(* CODESYS project RobotLibrary.library
   Company: Thorsten Brach
   Description: SRCI Robot Library
   Version: 1.5.7.0
   Placeholder: RobotLibrary
   Author: Thorsten Brach
   Title: RobotLibrary

Project tree, tasks and I/O mapping:
  libraries: RobotLibrarySysDep, * (Thorsten Brach); Tc2_Standard, 3.4.5.0 (Beckhoff Automation GmbH)
  Library/
    Constants/
      global variables RobotLibraryConstants
      global variables RobotLibraryDefines
    Enumerations/
      ArmConfig/
        data type ArmConfigElbow
        data type ArmConfigShoulder
        data type ArmConfigWrist
      Events/
        data type RobotLibraryErrorIdEnum
        data type RobotLibraryInfoIdEnum
        data type RobotLibraryWarningIdEnum
      Flag/
        data type SequenceFlag
        data type SequenceFlagEnum
      Level/
        data type LogLevel
        data type LogLevelEnum
        data type MessageLevel
        data type MessageLevelEnum
        data type PriorityLevel
      Miscellaneous/
        data type AxisUnit
        data type CircPlane
        data type ComDirection
        data type ControlHalfByte
        data type ErrorReaction
        data type LoadMeasurementSteps
        data type PathChoice
        data type ReferenceElement
        data type Severity
        data type SyncDirection
        data type SyncReaction
        data type SyncTime
        data type TriggerCondition
        data type UnitLimitAxis
      Mode/
        data type AbortingMode
        data type AbortingModeEnum
        data type BlendingMode
        data type CircMode
        data type CollisionReactionMode
        data type ConnectionMode
        data type DefinitionMode
        data type DetectionMode
        data type ErrorTriggerMode
        data type ExecutionMode
        data type FrameCalculationMode
        data type FunctionMode
        data type InterpolationMode
        data type JogMode
        data type LimitMode
        data type LoadMeasurementMode
        data type LogonMode
        data type MeasuringIoMode
        data type MeasuringUnitMode
        data type OperationMode
        data type OrientationMode
        data type OriMode
        data type ProcessingMode
        data type ProcessingModeEnum
        data type ResistanceForceMode
        data type ReturnMode
        data type SensorConnectionMode
        data type SingularityAvoidanceMode
        data type SplineMode
        data type StepMode
        data type StopMode
        data type SyncInMode
        data type SyncMode
        data type ThresholdMode
        data type ToolCalculationMode
        data type TrajectoryMode
        data type TransformMode
        data type TriggerModeIo
        data type TriggerModeLimit
        data type TriggerModeMeasurement
        data type TriggerReactionMode
        data type TurnMode
        data type WorkAreaReactionMode
      State/
        data type ActiveCommandRegisterState
        data type BufferStateCmd
        data type BufferStateRsp
        data type CmdMessageState
        data type InitializationState
        data type RaPowerState
        data type RaSequenceState
        data type RiState
        data type TelegramState
      Type/
        data type AreaType
        data type AreaTypeEnum
        data type AxesGroupParameterCmdEntries
        data type CmdType
        data type ConveyorType
        data type DataType
        data type MessageType
        data type ReferenceType
        data type UnitType
    Functions/
      Check/
        function IsDefaultDynamicsEqual [ST]
        function IsFrameDataEqual [ST]
        function IsLoadDataEqual [ST]
        function IsReferenceDynamicsEqual [ST]
        function IsSwLimitsEqual [ST]
        function IsToolDataEqual [ST]
        function IsWorkAreaEqual [ST]
      Common/
        function CheckTimeout [ST]
        function SetTimeout [ST]
      Convert/
        DT/
          function DATE_TO_IEC_DATE [ST]
          function IEC_DATE_TO_DATE [ST]
          function IEC_TIME_TO_TIME [ST]
          function IEC_TIMESTAMP_TO_DT [ST]
          function IEC_TIMESTAMP_TO_SYSTEMTIME [ST]
          function SYSTEMTIME_TO_IEC_TIMESTAMP [ST]
          function TIME_TO_IEC_TIME [ST]
        Misc/
          function ArmConfigParameterToBytes [ST]
          function BytesToRCSupportedFunctions [ST]
          function ByteToAxisExternalUnit [ST]
          function ByteToAxisExternalUsed [ST]
          function ByteToAxisJointUnit [ST]
          function ByteToAxisJointUsed [ST]
          function ByteToFragmentAction [ST]
          function ByteToVersion [ST]
          function CombineBytesToUint [ST]
          function CombineHalfBytes [ST]
          function CombineHalfSints [ST]
          function DwordToRaStatusWord [ST]
          function FragmentActionToByte [ST]
          function PERCENT_INT_TO_REAL [ST]
          function PERCENT_UINT_TO_REAL [ST]
          function PlcOptionalCyclicToUint [ST]
          function REAL_TO_PERCENT_INT [ST]
          function REAL_TO_PERCENT_UINT [ST]
          function RobOptionalCyclicToUint [ST]
          function SIGN_MAGNITUDE_TO_TURN [ST]
          function SyncModesToDataEnableSync [ST]
          function TURN_TO_SIGN_MAGNITUDE [ST]
          function VersionToByte [ST]
          function WordToArmConfigElbow [ST]
          function WordToArmConfigShoulder [ST]
          function WordToArmConfigWrist [ST]
        TO_STRING/
          function ABORTING_MODE_TO_STRING [ST]
          function ALARM_MESSAGE_TO_STRING [ST]
          function AREA_TYPE_TO_STRING [ST]
          function ARM_CONFIG_ELBOW_TO_STRING [ST]
          function ARM_CONFIG_SHOULDER_TO_STRING [ST]
          function ARM_CONFIG_TO_STRING [ST]
          function ARM_CONFIG_WRIST_TO_STRING [ST]
          function BLENDING_MODE_TO_STRING [ST]
          function BYTE_TO_STRING_BIN [ST]
          function CIRC_MODE_TO_STRING [ST]
          function CIRC_PLANE_TO_STRING [ST]
          function CMD_MESSAGE_STATE_TO_STRING [ST]
          function CMD_TYPE_TO_STRING [ST]
          function COLLISION_REACTION_MODE_TO_STRING [ST]
          function CONNECTION_MODE_TO_STRING [ST]
          function CONVEYOR_TYPE_TO_STRING [ST]
          function DATA_ENABLE_SYNC_TO_STRING [ST]
          function DATA_IN_SYNC_TO_STRING [ST]
          function DATA_TYPE_TO_STRING [ST]
          function DEFINITION_MODE_TO_STRING [ST]
          function DETECTION_MODE_TO_STRING [ST]
          function ERROR_REACTION_TO_STRING [ST]
          function ERROR_TRIGGER_MODE_TO_STRING [ST]
          function EXECUTION_MODE_TO_STRING [ST]
          function EXTERNAL_AXES_FLAGS_TO_STRING [ST]
          function FRAGMENT_ACTION_TO_STRING [ST]
          function FRAME_CALCULATION_MODE_TO_STRING [ST]
          function IEC_DATE_TO_STRING [ST]
          function IEC_TIME_TO_STRING [ST]
          function INTERPOLATION_MODE_TO_STRING [ST]
          function JOG_CONTROL_TO_STRING [ST]
          function JOG_MODE_TO_STRING [ST]
          function LIMIT_MODE_TO_STRING [ST]
          function LOAD_MEASUREMENT_MODE_TO_STRING [ST]
          function LOAD_MEASUREMENT_STEPS_TO_STRING [ST]
          function LOG_LEVEL_TO_STRING [ST]
          function LOGON_MODE_TO_STRING [ST]
          function MEASUREING_UNIT_MODE_TO_STRING [ST]
          function MEASURING_IO_MODE_TO_STRING [ST]
          function MEASURING_UNIT_MODE_TO_STRING [ST]
          function MESSAGE_CODE_TO_STRING [ST]
          function MESSAGE_LEVEL_TO_STRING [ST]
          function MESSAGE_TYPE_TO_STRING [ST]
          function OPERATION_MODE_TO_STRING [ST]
          function ORI_MODE_TO_STRING [ST]
          function PATH_CHOICE_TO_STRING [ST]
          function PROCESSING_MODE_TO_STRING [ST]
          function REFERENCE_ELEMENT_TO_STRING [ST]
          function REFERENCE_TYPE_TO_STRING [ST]
          function RESISTANT_FORCE_MODE_TO_STRING [ST]
          function RETURN_MODE_TO_STRING [ST]
          function ROBOT_AXES_FLAGS_TO_STRING [ST]
          function SENSOR_CONNECTION_MODE_TO_STRING [ST]
          function SEQUENCE_FLAG_TO_STRING [ST]
          function SEVERITY_TO_STRING [ST]
          function SINGULARITY_AVOIDANCE_MODE_TO_STRING [ST]
          function SPLINE_MODE_TO_STRING [ST]
          function STEP_MODE_TO_STRING [ST]
          function STOP_MODE_TO_STRING [ST]
          function SYNC_IN_MODE_TO_STRING [ST]
          function SYNC_MODE_TO_STRING [ST]
          function SYNC_REACTION_TO_STRING [ST]
          function SYNC_TIME_TO_STRING [ST]
          function TELEGRAM_CONTROL_TO_STRING [ST]
          function TELEGRAM_STATE_TO_STRING [ST]
          function THRESHOLD_MODE_TO_STRING [ST]
          function TOOL_CALCULATION_MODE_TO_STRING [ST]
          function TRAJECTORY_MODE_TO_STRING [ST]
          function TRANSFORM_MODE_TO_STRING [ST]
          function TRIGGER_CONDITION_TO_STRING [ST]
          function TRIGGER_MODE_IO_TO_STRING [ST]
          function TRIGGER_MODE_LIMIT_TO_STRING [ST]
          function TRIGGER_MODE_MEASUREMENT_TO_STRING [ST]
          function TRIGGER_REACTION_MODE_TO_STRING [ST]
          function TURN_MODE_TO_STRING [ST]
          function UNIT_LIMIT_AXIS_TO_STRING [ST]
          function VALID_REAL_TO_STRING [ST]
          function WORD_TO_STRING_BIN [ST]
          function WORD_TO_STRING_HEX [ST]
          function WORK_AREA_REACTION_MODE_TO_STRING [ST]
      String/
        function StrPadRight [ST]
        function StrReplace [ST]
      Swap/
        function GetHalfeByteHi [ST]
        function GetHalfeByteLo [ST]
        function SwapBytes [ST]
        function SwapDword [ST]
        function SwapIecDate [ST]
        function SwapIecTime [ST]
        function SwapInt [ST]
        function SwapReal [ST]
        function SwapUdint [ST]
        function SwapUint [ST]
        function SwapWord [ST]
    Interfaces/
      interface IMessageLogger: AddMessageLog, AddSystemLog
      interface IRobotLibraryCommandFB: CallBack, CommandData
    Parameter/
      global variables RobotLibraryParameter
    POUs/
      _internal/
        BaseFBs/
          function block RobotLibraryBaseEnableFB [ST]: OnCall, OnExecCancel, OnExecErrorClear, OnExecRun, OnExecStart, OnUpdateStateFlags, Reset
          function block RobotLibraryBaseExecuteFB [ST]: OnCall, OnExecCancel, OnExecErrorClear, OnExecRun, OnExecStart, OnUpdateStateFlags, Reset
          function block RobotLibraryBaseFB [ST]: CallBack, CheckFunctionSupported, CheckParameterChanged, CheckParameterValid, CreateCommandPayload, HasError, HasInfo, HasWarning, OnApplyOutCmd, OnCall, OnExecRun, OnOnlineChange, OnUpdateStateFlags, ParseResponsePayload, Reset, SetError, SetInfo, SetWarning
          function block RobotLibraryLogFB [ST]: CreateLogMessage, CreateLogMessagePara1, CreateLogMessagePara2, CreateLogMessagePara3, CreateLogMessagePara4, CreateLogMessagePara5, CreateLogMessagePara6, MyType
        LogFBs/
          function block AxesGroupMessageLogFB [ST]: AddMessageLog, AddMessageLogByParameter, AddSystemLog, CheckMessageCodePresent, DeleteMessages, DeleteSystemLogs
        Recv/
          function block RobotLibraryRecvDataBaseFB [ST]: GetArmConfig, GetBool, GetByte, GetDataBlock, GetDataInSync, GetDword, GetFragmentAction, GetHalfeByte1, GetHalfeByte2, GetIecDate, GetIecTime, GetInt, GetReal, GetSint, GetString, GetTrackingStatus, GetTurnNumbers, GetUdint, GetUint, GetUsint, GetWord, Reset, UpdatePointer
          function block RobotLibraryRecvDataFB [ST]: GetLifeSignFooter, UpdatePointer
          function block RobotLibraryResponseDataFB [ST]: IsPayloadRemaining, Reset, UpdatePointer
        Send/
          function block RobotLibraryCommandDataFB [ST]: Reset, UpdatePointer
          function block RobotLibrarySendDataBaseFB [ST]: AddArmConfig, AddBool, AddByte, AddDataBlock, AddDataEnableSync, AddDataInSync, AddDword, AddHalfBytes, AddIecDate, AddIecTime, AddInt, AddReal, AddSint, AddString, AddTime, AddTurnNumber, AddUdint, AddUint, AddUsint, Reset, UpdatePointer
          function block RobotLibrarySendDataFB [ST]: Reset, SetLifeSignFooter, UpdatePointer
        SystemData/
          function block AxesGroupSystemDataFB [ST]: UpdateDefaultDynamics, UpdateFrameData, UpdateLoadData, UpdateReferenceDynamics, UpdateSWLimits, UpdateToolData, UpdateWorAreas
        function block ActiveCommandRegisterFB [ST]: AddCmd, AddRsp, FB_init, ManageRegister, NotifyParameterChanged, OnOnlineChange, RemoveCmd, Reset, UpdateExecutionOrderList
      Additional/
        MC_AbortMeasuringInput/
          Structures/
            data type AbortMeasuringInputOutCmd
            data type AbortMeasuringInputParCmd
            data type AbortMeasuringInputRecvData
            data type AbortMeasuringInputSendData
          function block MC_AbortMeasuringInputFB [ST]: CheckAddParameter, CheckFunctionSupported, CheckParameterChanged, CheckParameterValid, CreateCommandPayload, CreateCommandPayloadLog, FB_init, OnExecRun, OnUpdateStateFlags, ParseResponsePayload, ParseResponsePayloadLog, Reset
        MC_ActivateNextCommand/
          Structures/
            data type ActivateNextCommandOutCmd
            data type ActivateNextCommandParCmd
            data type ActivateNextCommandRecvData
            data type ActivateNextCommandSendData
          function block MC_ActivateNextCommandFB [ST]: CheckAddParameter, CheckFunctionSupported, CheckParameterChanged, CheckParameterValid, CreateCommandPayload, CreateCommandPayloadLog, FB_init, OnApplyOutCmd, OnExecRun, OnUpdateStateFlags, ParseResponsePayload, ParseResponsePayloadLog, Reset
        MC_AvoidSingularity/
          Structures/
            data type AvoidSingularityOutCmd
            data type AvoidSingularityParCmd
            data type AvoidSingularityRecvData
            data type AvoidSingularitySendData
          function block MC_AvoidSingularityFB [ST]: CheckAddParameter, CheckFunctionSupported, CheckParameterChanged, CheckParameterValid, CreateCommandPayload, CreateCommandPayloadLog, FB_init, OnExecCancel, OnExecErrorClear, OnExecRun, OnUpdateStateFlags, ParseResponsePayload, ParseResponsePayloadLog, Reset
        MC_BrakeTest/
          Structures/
            data type BrakeTestOutCmd
            data type BrakeTestParCmd
            data type BrakeTestRecvData
            data type BrakeTestSendData
          function block MC_BrakeTestFB [ST]: CheckAddParameter, CheckFunctionSupported, CheckParameterChanged, CheckParameterValid, CreateCommandPayload, CreateCommandPayloadLog, FB_init, OnApplyOutCmd, OnExecRun, OnUpdateStateFlags, ParseResponsePayload, ParseResponsePayloadLog, Reset
        MC_CallSubprogram/
          Structures/
            data type CallSubprogramOutCmd
            data type CallSubprogramParCmd
            data type CallSubprogramRecvData
            data type CallSubprogramSendData
          function block MC_CallSubprogramFB [ST]: CheckAddParameter, CheckFunctionSupported, CheckParameterChanged, CheckParameterValid, CreateCommandPayload, CreateCommandPayloadLog, FB_init, OnApplyOutCmd, OnExecRun, OnUpdateStateFlags, ParseResponsePayload, ParseResponsePayloadLog, Reset
        MC_CollisionDetection/
          Structures/
            data type CollisionDetectionOutCmd
            data type CollisionDetectionParCmd
            data type CollisionDetectionRecvData
            data type CollisionDetectionSendData
          function block MC_CollisionDetectionFB [ST]: CheckAddParameter, CheckFunctionSupported, CheckParameterChanged, CheckParameterValid, CreateCommandPayload, CreateCommandPayloadLog, FB_init, OnExecRun, OnUpdateStateFlags, ParseResponsePayload, ParseResponsePayloadLog, Reset
        MC_ExchangeConfiguration/
          Structures/
            data type ExchangeConfigurationOutCmd
            data type ExchangeConfigurationParCmd
            data type ExchangeConfigurationRecvData
            data type ExchangeConfigurationSendData
          function block MC_ExchangeConfigurationFB [ST]: CheckAddParameter, CheckFunctionSupported, CheckParameterChanged, CheckParameterValid, CreateCommandPayload, CreateCommandPayloadLog, FB_init, OnApplyOutCmd, OnExecCancel, OnExecErrorClear, OnExecRun, OnUpdateStateFlags, ParseResponsePayload, ParseResponsePayloadLog, Reset
        MC_FreeDrive/
          Structures/
            data type FreeDriveOutCmd
            data type FreeDriveParCmd
            data type FreeDriveRecvData
            data type FreeDriveSendData
          function block MC_FreeDriveFB [ST]: CheckAddParameter, CheckFunctionSupported, CheckParameterChanged, CreateCommandPayload, CreateCommandPayloadLog, FB_init, OnExecCancel, OnExecErrorClear, OnExecRun, OnUpdateStateFlags, ParseResponsePayload, ParseResponsePayloadLog, Reset
        MC_MeasuringInput/
          Structures/
            data type MeasuringInputOutCmd
            data type MeasuringInputParCmd
            data type MeasuringInputRecvData
            data type MeasuringInputSendData
          function block MC_MeasuringInputFB [ST]: CheckAddParameter, CheckFunctionSupported, CheckParameterChanged, CheckParameterValid, CreateCommandPayload, CreateCommandPayloadLog, FB_init, OnApplyOutCmd, OnExecRun, OnUpdateStateFlags, ParseResponsePayload, ParseResponsePayloadLog, Reset
        MC_OpenBrake/
          Structures/
            data type OpenBrakeOutCmd
            data type OpenBrakeParCmd
            data type OpenBrakeRecvData
            data type OpenBrakeSendData
          function block MC_OpenBrakeFB [ST]: CheckAddParameter, CheckFunctionSupported, CheckParameterChanged, CheckParameterValid, CreateCommandPayload, CreateCommandPayloadLog, FB_init, OnApplyOutCmd, OnExecCancel, OnExecErrorClear, OnExecRun, OnUpdateStateFlags, ParseResponsePayload, ParseResponsePayloadLog, Reset
        MC_PathAccuracyMode/
          Structures/
            data type PathAccuracyModeOutCmd
            data type PathAccuracyModeParCmd
            data type PathAccuracyModeRecvData
            data type PathAccuracyModeSendData
          function block MC_PathAccuracyModeFB [ST]: CheckAddParameter, CheckFunctionSupported, CheckParameterChanged, CreateCommandPayload, CreateCommandPayloadLog, FB_init, OnExecCancel, OnExecErrorClear, OnExecRun, OnUpdateStateFlags, ParseResponsePayload, ParseResponsePayloadLog, Reset
        MC_ReadCallSubprogramCyclic/
          Structures/
            data type ReadCallSubprogramCyclicOutCmd
            data type ReadCallSubprogramCyclicParCmd
          function block MC_ReadCallSubprogramCyclicFB [ST]: CheckFunctionSupported, CheckParameterChanged, CheckParameterValid, CreateCommandParameterLog, FB_init, OnExecErrorClear, OnExecRun, Reset
        MC_ReadSafeReferencePosition/
          Structures/
            data type ReadSafeReferencePositionOutCmd
            data type ReadSafeReferencePositionParCmd
            data type ReadSafeReferencePositionRecvData
            data type ReadSafeReferencePositionSendData
          function block MC_ReadSafeReferencePositionFB [ST]: CheckAddParameter, CheckFunctionSupported, CheckParameterChanged, CheckParameterValid, CreateCommandPayload, CreateCommandPayloadLog, FB_init, OnApplyOutCmd, OnExecRun, OnUpdateStateFlags, ParseResponsePayload, ParseResponsePayloadLog, Reset
        MC_SafeReferencing/
          Structures/
            data type SafeReferencingOutCmd
            data type SafeReferencingParCmd
            data type SafeReferencingRecvData
            data type SafeReferencingSendData
          function block MC_SafeReferencingFB [ST]: CheckAddParameter, CheckFunctionSupported, CheckParameterChanged, CheckParameterValid, CreateCommandPayload, CreateCommandPayloadLog, FB_init, OnApplyOutCmd, OnExecRun, OnUpdateStateFlags, ParseResponsePayload, ParseResponsePayloadLog, Reset
        MC_ShiftPosition/
          Structures/
            data type ShiftPositionOutCmd
            data type ShiftPositionParCmd
            data type ShiftPositionRecvData
            data type ShiftPositionSendData
          function block MC_ShiftPositionFB [ST]: CheckAddParameter, CheckFunctionSupported, CheckParameterChanged, CheckParameterValid, CreateCommandPayload, CreateCommandPayloadLog, FB_init, OnApplyOutCmd, OnExecRun, OnUpdateStateFlags, ParseResponsePayload, ParseResponsePayloadLog, Reset
        MC_SoftSwitchTcp/
          Structures/
            data type SoftSwitchTcpOutCmd
            data type SoftSwitchTcpParCmd
            data type SoftSwitchTcpRecvData
            data type SoftSwitchTcpSendData
          function block MC_SoftSwitchTcpFB [ST]: CheckAddParameter, CheckFunctionSupported, CheckParameterChanged, CheckParameterValid, CreateCommandPayload, CreateCommandPayloadLog, FB_init, OnApplyOutCmd, OnExecRun, OnUpdateStateFlags, ParseResponsePayload, ParseResponsePayloadLog, Reset
        MC_StopSubprogram/
          Structures/
            data type StopSubprogramOutCmd
            data type StopSubprogramParCmd
            data type StopSubprogramRecvData
            data type StopSubprogramSendData
          function block MC_StopSubprogramFB [ST]: CheckAddParameter, CheckFunctionSupported, CheckParameterChanged, CheckParameterValid, CreateCommandPayload, CreateCommandPayloadLog, FB_init, OnApplyOutCmd, OnExecRun, OnUpdateStateFlags, ParseResponsePayload, ParseResponsePayloadLog, Reset
        MC_UnitMeasurement/
          Structures/
            data type UnitMeasurementOutCmd
            data type UnitMeasurementParCmd
            data type UnitMeasurementRecvData
            data type UnitMeasurementSendData
          function block MC_UnitMeasurementFB [ST]: CheckAddParameter, CheckFunctionSupported, CheckParameterChanged, CheckParameterValid, CreateCommandPayload, CreateCommandPayloadLog, FB_init, OnApplyOutCmd, OnExecCancel, OnExecErrorClear, OnExecRun, OnUpdateStateFlags, ParseResponsePayload, ParseResponsePayloadLog, Reset
        MC_WriteCallSubprogramCyclic/
          Structures/
            data type WriteCallSubprogramCyclicOutCmd
            data type WriteCallSubprogramCyclicParCmd
          function block MC_WriteCallSubprogramCyclicFB [ST]: CheckFunctionSupported, FB_init, OnExecErrorClear, OnExecRun
      AdvancedMove/
        MC_MoveApproachDirect/
          Structures/
            data type MoveApproachDirectOutCmd
            data type MoveApproachDirectParCmd
            data type MoveApproachDirectRecvData
            data type MoveApproachDirectSendData
          function block MC_MoveApproachDirectFB [ST]: CheckAddParameter, CheckFunctionSupported, CheckParameterChanged, CheckParameterValid, CreateCommandPayload, CreateCommandPayloadLog, FB_init, OnApplyOutCmd, OnExecRun, OnUpdateStateFlags, ParseResponsePayload, ParseResponsePayloadLog, Reset
        MC_MoveApproachLinear/
          Structures/
            data type MoveApproachLinearOutCmd
            data type MoveApproachLinearParCmd
            data type MoveApproachLinearRecvData
            data type MoveApproachLinearSendData
          function block MC_MoveApproachLinearFB [ST]: CheckAddParameter, CheckFunctionSupported, CheckParameterChanged, CheckParameterValid, CreateCommandPayload, CreateCommandPayloadLog, FB_init, OnApplyOutCmd, OnExecRun, OnUpdateStateFlags, ParseResponsePayload, ParseResponsePayloadLog, Reset
        MC_MoveAxesRelative/
          Structures/
            data type MoveAxesRelativeOutCmd
            data type MoveAxesRelativeParCmd
            data type MoveAxesRelativeRecvData
            data type MoveAxesRelativeSendData
          function block MC_MoveAxesRelativeFB [ST]: CheckAddParameter, CheckFunctionSupported, CheckParameterChanged, CheckParameterValid, CreateCommandPayload, CreateCommandPayloadLog, FB_init, OnApplyOutCmd, OnExecRun, OnUpdateStateFlags, ParseResponsePayload, ParseResponsePayloadLog, Reset
        MC_MoveCircularAbsolute/
          Structures/
            data type MoveCircularAbsoluteOutCmd
            data type MoveCircularAbsoluteParCmd
            data type MoveCircularAbsoluteRecvData
            data type MoveCircularAbsoluteSendData
          function block MC_MoveCircularAbsoluteFB [ST]: CheckAddParameter, CheckFunctionSupported, CheckParameterChanged, CheckParameterValid, CreateCommandPayload, CreateCommandPayloadLog, FB_init, OnApplyOutCmd, OnExecRun, OnUpdateStateFlags, ParseResponsePayload, ParseResponsePayloadLog, Reset
        MC_MoveCircularCamFB/
          Structures/
            data type MoveCircularCamOutCmd
            data type MoveCircularCamParCmd
            data type MoveCircularCamRecvData
            data type MoveCircularCamSendData
          function block MC_MoveCircularCamFB [ST]: CheckAddParameter, CheckFunctionSupported, CheckParameterChanged, CheckParameterValid, CreateCommandPayload, CreateCommandPayloadLog, FB_init, OnApplyOutCmd, OnExecRun, OnUpdateStateFlags, ParseResponsePayload, ParseResponsePayloadLog, Reset
        MC_MoveCircularRelative/
          Structures/
            data type MoveCircularRelativeOutCmd
            data type MoveCircularRelativeParCmd
            data type MoveCircularRelativeRecvData
            data type MoveCircularRelativeSendData
          function block MC_MoveCircularRelativeFB [ST]: CheckAddParameter, CheckFunctionSupported, CheckParameterChanged, CheckParameterValid, CreateCommandPayload, CreateCommandPayloadLog, FB_init, OnApplyOutCmd, OnExecRun, OnUpdateStateFlags, ParseResponsePayload, ParseResponsePayloadLog, Reset
        MC_MoveDepartDirect/
          Structures/
            data type MoveDepartDirectOutCmd
            data type MoveDepartDirectParCmd
            data type MoveDepartDirectRecvData
            data type MoveDepartDirectSendData
          function block MC_MoveDepartDirectFB [ST]: CheckAddParameter, CheckFunctionSupported, CheckParameterChanged, CheckParameterValid, CreateCommandPayload, CreateCommandPayloadLog, FB_init, OnApplyOutCmd, OnExecRun, OnUpdateStateFlags, ParseResponsePayload, ParseResponsePayloadLog, Reset
        MC_MoveDepartLinear/
          Structures/
            data type MoveDepartLinearOutCmd
            data type MoveDepartLinearParCmd
            data type MoveDepartLinearRecvData
            data type MoveDepartLinearSendData
          function block MC_MoveDepartLinearFB [ST]: CheckAddParameter, CheckFunctionSupported, CheckParameterChanged, CheckParameterValid, CreateCommandPayload, CreateCommandPayloadLog, FB_init, OnApplyOutCmd, OnExecRun, OnUpdateStateFlags, ParseResponsePayload, ParseResponsePayloadLog, Reset
        MC_MoveDirectCam/
          Structures/
            data type MoveDirectCamOutCmd
            data type MoveDirectCamParCmd
            data type MoveDirectCamRecvData
            data type MoveDirectCamSendData
          function block MC_MoveDirectCamFB [ST]: CheckAddParameter, CheckFunctionSupported, CheckParameterChanged, CheckParameterValid, CreateCommandPayload, CreateCommandPayloadLog, FB_init, OnApplyOutCmd, OnExecRun, OnUpdateStateFlags, ParseResponsePayload, ParseResponsePayloadLog, Reset
        MC_MoveDirectOffset/
          Structures/
            data type MoveDirectOffsetOutCmd
            data type MoveDirectOffsetParCmd
            data type MoveDirectOffsetRecvData
            data type MoveDirectOffsetSendData
          function block MC_MoveDirectOffsetFB [ST]: CheckAddParameter, CheckFunctionSupported, CheckParameterChanged, CheckParameterValid, CreateCommandPayload, CreateCommandPayloadLog, FB_init, OnApplyOutCmd, OnExecRun, OnUpdateStateFlags, ParseResponsePayload, ParseResponsePayloadLog, Reset
        MC_MoveDirectRelative/
          Structures/
            data type MoveDirectRelativeOutCmd
            data type MoveDirectRelativeParCmd
            data type MoveDirectRelativeRecvData
            data type MoveDirectRelativeSendData
          function block MC_MoveDirectRelativeFB [ST]: CheckAddParameter, CheckFunctionSupported, CheckParameterChanged, CheckParameterValid, CreateCommandPayload, CreateCommandPayloadLog, FB_init, OnApplyOutCmd, OnExecRun, OnUpdateStateFlags, ParseResponsePayload, ParseResponsePayloadLog, Reset
        MC_MoveLinearAbsoluteJ/
          Structures/
            data type MoveLinearAbsoluteJOutCmd
            data type MoveLinearAbsoluteJParCmd
            data type MoveLinearAbsoluteJRecvData
            data type MoveLinearAbsoluteJSendData
          function block MC_MoveLinearAbsoluteJFB [ST]: CheckAddParameter, CheckFunctionSupported, CheckParameterChanged, CheckParameterValid, CreateCommandPayload, CreateCommandPayloadLog, FB_init, OnApplyOutCmd, OnExecRun, OnUpdateStateFlags, ParseResponsePayload, ParseResponsePayloadLog, Reset
        MC_MoveLinearCam/
          Structures/
            data type MoveLinearCamOutCmd
            data type MoveLinearCamParCmd
            data type MoveLinearCamRecvData
            data type MoveLinearCamSendData
          function block MC_MoveLinearCamFB [ST]: CheckAddParameter, CheckFunctionSupported, CheckParameterChanged, CheckParameterValid, CreateCommandPayload, CreateCommandPayloadLog, FB_init, OnApplyOutCmd, OnExecRun, OnUpdateStateFlags, ParseResponsePayload, ParseResponsePayloadLog, Reset
        MC_MoveLinearOffset/
          Structures/
            data type MoveLinearOffsetOutCmd
            data type MoveLinearOffsetParCmd
            data type MoveLinearOffsetRecvData
            data type MoveLinearOffsetSendData
          function block MC_MoveLinearOffsetFB [ST]: CheckAddParameter, CheckFunctionSupported, CheckParameterChanged, CheckParameterValid, CreateCommandPayload, CreateCommandPayloadLog, FB_init, OnApplyOutCmd, OnExecRun, OnUpdateStateFlags, ParseResponsePayload, ParseResponsePayloadLog, Reset
        MC_MoveLinearRelative/
          Structures/
            data type MoveLinearRelativeOutCmd
            data type MoveLinearRelativeParCmd
            data type MoveLinearRelativeRecvData
            data type MoveLinearRelativeSendData
          function block MC_MoveLinearRelativeFB [ST]: CheckAddParameter, CheckFunctionSupported, CheckParameterChanged, CheckParameterValid, CreateCommandPayload, CreateCommandPayloadLog, FB_init, OnApplyOutCmd, OnExecRun, OnUpdateStateFlags, ParseResponsePayload, ParseResponsePayloadLog, Reset
        MC_MovePickPlaceDirect/
          Structures/
            data type MovePickPlaceDirectOutCmd
            data type MovePickPlaceDirectParCmd
            data type MovePickPlaceDirectRecvData
            data type MovePickPlaceDirectSendData
          function block MC_MovePickPlaceDirectFB [ST]: CheckAddParameter, CheckFunctionSupported, CheckParameterChanged, CheckParameterValid, CreateCommandPayload, CreateCommandPayloadLog, FB_init, OnApplyOutCmd, OnExecRun, OnUpdateStateFlags, ParseResponsePayload, ParseResponsePayloadLog, Reset
        MC_MovePickPlaceLinear/
          Structures/
            data type MovePickPlaceLinearOutCmd
            data type MovePickPlaceLinearParCmd
            data type MovePickPlaceLinearRecvData
            data type MovePickPlaceLinearSendData
          function block MC_MovePickPlaceLinearFB [ST]: CheckAddParameter, CheckFunctionSupported, CheckParameterChanged, CheckParameterValid, CreateCommandPayload, CreateCommandPayloadLog, FB_init, OnApplyOutCmd, OnExecRun, OnUpdateStateFlags, ParseResponsePayload, ParseResponsePayloadLog, Reset
      BasicMove/
        MC_ChangeSpeedOverride/
          Structures/
            data type ChangeSpeedOverrideOutCmd
            data type ChangeSpeedOverrideParCmd
            data type ChangeSpeedOverrideRecvData
            data type ChangeSpeedOverrideSendData
          function block MC_ChangeSpeedOverrideFB [ST]: CheckAddParameter, CheckFunctionSupported, CheckParameterChanged, CheckParameterValid, CreateCommandPayload, CreateCommandPayloadLog, FB_init, OnExecRun, OnUpdateStateFlags, ParseResponsePayload, ParseResponsePayloadLog, Reset
        MC_GroupContinue/
          Structures/
            data type GroupContinueOutCmd
            data type GroupContinueParCmd
            data type GroupContinueRecvData
            data type GroupContinueSendData
          function block MC_GroupContinueFB [ST]: CheckAddParameter, CheckFunctionSupported, CheckParameterChanged, CheckSynchronizationValid, CreateCommandPayload, CreateCommandPayloadLog, FB_init, OnExecRun, OnUpdateStateFlags, ParseResponsePayload, ParseResponsePayloadLog, Reset
        MC_GroupInterrupt/
          Structures/
            data type GroupInterruptOutCmd
            data type GroupInterruptParCmd
            data type GroupInterruptRecvData
            data type GroupInterruptSendData
          function block MC_GroupInterruptFB [ST]: CheckAddParameter, CheckFunctionSupported, CheckParameterChanged, CreateCommandPayload, CreateCommandPayloadLog, FB_init, OnExecRun, OnUpdateStateFlags, ParseResponsePayload, ParseResponsePayloadLog, Reset
        MC_GroupJog/
          Structures/
            data type GroupJogOutCmd
            data type GroupJogParCmd
            data type GroupJogRecvData
            data type GroupJogSendData
          function block MC_GroupJogFB [ST]: CheckAddParameter, CheckFunctionSupported, CheckParameterChanged, CheckParameterValid, CreateCommandPayload, CreateCommandPayloadLog, FB_init, OnApplyOutCmd, OnExecCancel, OnExecErrorClear, OnExecRun, OnUpdateStateFlags, ParseResponsePayload, ParseResponsePayloadLog, Reset
        MC_GroupStop/
          Structures/
            data type GroupStopOutCmd
            data type GroupStopParCmd
            data type GroupStopRecvData
            data type GroupStopSendData
          function block MC_GroupStopFB [ST]: CheckAddParameter, CheckFunctionSupported, CheckParameterChanged, CreateCommandPayload, CreateCommandPayloadLog, FB_init, OnExecRun, OnUpdateStateFlags, ParseResponsePayload, ParseResponsePayloadLog, Reset
        MC_MoveAxesAbsolute/
          Structures/
            data type MoveAxesAbsoluteOutCmd
            data type MoveAxesAbsoluteParCmd
            data type MoveAxesAbsoluteRecvData
            data type MoveAxesAbsoluteSendData
          function block MC_MoveAxesAbsoluteFB [ST]: CheckAddParameter, CheckFunctionSupported, CheckParameterChanged, CheckParameterValid, CreateCommandPayload, CreateCommandPayloadLog, FB_init, OnApplyOutCmd, OnExecRun, OnUpdateStateFlags, ParseResponsePayload, ParseResponsePayloadLog, Reset
        MC_MoveDirectAbsolute/
          Structures/
            data type MoveDirectAbsoluteOutCmd
            data type MoveDirectAbsoluteParCmd
            data type MoveDirectAbsoluteRecvData
            data type MoveDirectAbsoluteSendData
          function block MC_MoveDirectAbsoluteFB [ST]: CheckAddParameter, CheckFunctionSupported, CheckParameterChanged, CheckParameterValid, CreateCommandPayload, CreateCommandPayloadLog, FB_init, OnApplyOutCmd, OnExecRun, OnUpdateStateFlags, ParseResponsePayload, ParseResponsePayloadLog, Reset
        MC_MoveLinearAbsolute/
          Structures/
            data type MoveLinearAbsoluteOutCmd
            data type MoveLinearAbsoluteParCmd
            data type MoveLinearAbsoluteRecvData
            data type MoveLinearAbsoluteSendData
          function block MC_MoveLinearAbsoluteFB [ST]: CheckAddParameter, CheckFunctionSupported, CheckParameterChanged, CheckParameterValid, CreateCommandPayload, CreateCommandPayloadLog, FB_init, OnApplyOutCmd, OnExecRun, OnUpdateStateFlags, ParseResponsePayload, ParseResponsePayloadLog, Reset
        MC_ReturnToPrimary/
          Structures/
            data type ReturnToPrimaryOutCmd
            data type ReturnToPrimaryParCmd
            data type ReturnToPrimaryRecvData
            data type ReturnToPrimarySendData
          function block MC_ReturnToPrimaryFB [ST]: CheckAddParameter, CheckFunctionSupported, CheckParameterChanged, CheckParameterValid, CreateCommandPayload, CreateCommandPayloadLog, FB_init, OnApplyOutCmd, OnExecRun, OnUpdateStateFlags, ParseResponsePayload, ParseResponsePayloadLog, Reset
      Calculation/
        MC_CalculateCartesianPosition/
          Structures/
            data type CalculateCartesianPositionOutCmd
            data type CalculateCartesianPositionParCmd
            data type CalculateCartesianPositionRecvData
            data type CalculateCartesianPositionSendData
          function block MC_CalculateCartesianPositionFB [ST]: CheckAddParameter, CheckFunctionSupported, CheckParameterChanged, CheckParameterValid, CreateCommandPayload, CreateCommandPayloadLog, FB_init, OnApplyOutCmd, OnExecRun, OnUpdateStateFlags, ParseResponsePayload, ParseResponsePayloadLog, Reset
        MC_CalculateForwardKinematic/
          Structures/
            data type CalculateForwardKinematicOutCmd
            data type CalculateForwardKinematicParCmd
            data type CalculateForwardKinematicRecvData
            data type CalculateForwardKinematicSendData
          function block MC_CalculateForwardKinematicFB [ST]: CheckAddParameter, CheckFunctionSupported, CheckParameterChanged, CheckParameterValid, CreateCommandPayload, CreateCommandPayloadLog, FB_init, OnApplyOutCmd, OnExecRun, OnUpdateStateFlags, ParseResponsePayload, ParseResponsePayloadLog, Reset
        MC_CalculateFrame/
          Structures/
            data type CalculateFrameOutCmd
            data type CalculateFrameParCmd
            data type CalculateFrameRecvData
            data type CalculateFrameSendData
          function block MC_CalculateFrameFB [ST]: CheckAddParameter, CheckFunctionSupported, CheckParameterChanged, CheckParameterValid, CreateCommandPayload, CreateCommandPayloadLog, FB_init, OnApplyOutCmd, OnExecRun, OnUpdateStateFlags, ParseResponsePayload, ParseResponsePayloadLog, Reset
        MC_CalculateInverseKinematic/
          Structures/
            data type CalculateInverseKinematicOutCmd
            data type CalculateInverseKinematicParCmd
            data type CalculateInverseKinematicRecvData
            data type CalculateInverseKinematicSendData
          function block MC_CalculateInverseKinematicFB [ST]: CheckAddParameter, CheckFunctionSupported, CheckParameterChanged, CheckParameterValid, CreateCommandPayload, CreateCommandPayloadLog, FB_init, OnApplyOutCmd, OnExecRun, OnUpdateStateFlags, ParseResponsePayload, ParseResponsePayloadLog, Reset
        MC_CalculateTool/
          Structures/
            data type CalculateToolOutCmd
            data type CalculateToolParCmd
            data type CalculateToolRecvData
            data type CalculateToolSendData
          function block MC_CalculateToolFB [ST]: CheckAddParameter, CheckFunctionSupported, CheckParameterChanged, CheckParameterValid, CreateCommandPayload, CreateCommandPayloadLog, FB_init, OnApplyOutCmd, OnExecRun, OnUpdateStateFlags, ParseResponsePayload, ParseResponsePayloadLog, Reset
        MC_LoadMeasurementAutomatic/
          Structures/
            data type LoadMeasurementAutomaticOutCmd
            data type LoadMeasurementAutomaticParCmd
            data type LoadMeasurementAutomaticRecvData
            data type LoadMeasurementAutomaticSendData
          function block MC_LoadMeasurementAutomaticFB [ST]: CheckAddParameter, CheckFunctionSupported, CheckParameterChanged, CheckParameterValid, CreateCommandPayload, CreateCommandPayloadLog, FB_init, OnApplyOutCmd, OnExecRun, OnUpdateStateFlags, ParseResponsePayload, ParseResponsePayloadLog, Reset
        MC_LoadMeasurementSequential/
          Structures/
            data type LoadMeasurementSequentialOutCmd
            data type LoadMeasurementSequentialParCmd
            data type LoadMeasurementSequentialRecvData
            data type LoadMeasurementSequentialSendData
          function block MC_LoadMeasurementSequentialFB [ST]: CheckAddParameter, CheckFunctionSupported, CheckParameterChanged, CheckParameterValid, CreateCommandPayload, CreateCommandPayloadLog, FB_init, OnApplyOutCmd, OnExecRun, OnUpdateStateFlags, ParseResponsePayload, ParseResponsePayloadLog, Reset
      ConveyorTracking/
        MC_ActivateConveyorTracking/
          Structures/
            data type ActivateConveyorTrackingOutCmd
            data type ActivateConveyorTrackingParCmd
            data type ActivateConveyorTrackingRecvData
            data type ActivateConveyorTrackingSendData
          function block MC_ActivateConveyorTrackingFB [ST]: CheckAddParameter, CheckFunctionSupported, CheckParameterChanged, CheckParameterValid, CreateCommandPayload, CreateCommandPayloadLog, FB_init, OnApplyOutCmd, OnExecCancel, OnExecErrorClear, OnExecRun, OnUpdateStateFlags, ParseResponsePayload, ParseResponsePayloadLog, Reset
        MC_ConfigureConveyor/
          Structures/
            data type ConfigureConveyorOutCmd
            data type ConfigureConveyorParCmd
            data type ConfigureConveyorRecvData
            data type ConfigureConveyorSendData
          function block MC_ConfigureConveyorFB [ST]: CheckAddParameter, CheckFunctionSupported, CheckParameterChanged, CheckParameterValid, CreateCommandPayload, CreateCommandPayloadLog, FB_init, OnExecRun, OnUpdateStateFlags, ParseResponsePayload, ParseResponsePayloadLog, Reset
        MC_RedefineTrackingPos/
          Structures/
            data type RedefineTrackingPosOutCmd
            data type RedefineTrackingPosParCmd
            data type RedefineTrackingPosRecvData
            data type RedefineTrackingPosSendData
          function block MC_RedefineTrackingPosFB [ST]: CheckAddParameter, CheckFunctionSupported, CheckParameterChanged, CheckParameterValid, CreateCommandPayload, CreateCommandPayloadLog, FB_init, OnApplyOutCmd, OnExecRun, OnUpdateStateFlags, ParseResponsePayload, ParseResponsePayloadLog, Reset
        MC_SyncToConveyor/
          Structures/
            data type SyncToConveyorOutCmd
            data type SyncToConveyorParCmd
            data type SyncToConveyorRecvData
            data type SyncToConveyorSendData
          function block MC_SyncToConveyorFB [ST]: CheckAddParameter, CheckFunctionSupported, CheckParameterChanged, CheckParameterValid, CreateCommandPayload, CreateCommandPayloadLog, FB_init, OnApplyOutCmd, OnExecCancel, OnExecErrorClear, OnExecRun, OnUpdateStateFlags, ParseResponsePayload, ParseResponsePayloadLog, Reset
      ForceControl/
        MC_ForceControl/
          Structures/
            data type ForceControlOutCmd
            data type ForceControlParCmd
            data type ForceControlRecvData
            data type ForceControlSendData
          function block MC_ForceControlFB [ST]: CheckAddParameter, CheckFunctionSupported, CheckParameterChanged, CheckParameterValid, CreateCommandPayload, CreateCommandPayloadLog, FB_init, OnApplyOutCmd, OnExecCancel, OnExecErrorClear, OnExecRun, OnUpdateStateFlags, ParseResponsePayload, ParseResponsePayloadLog, Reset
        MC_ForceLimit/
          Structures/
            data type ForceLimitOutCmd
            data type ForceLimitParCmd
            data type ForceLimitRecvData
            data type ForceLimitSendData
          function block MC_ForceLimitFB [ST]: CheckAddParameter, CheckFunctionSupported, CheckParameterChanged, CheckParameterValid, CreateCommandPayload, CreateCommandPayloadLog, FB_init, OnApplyOutCmd, OnExecCancel, OnExecErrorClear, OnExecRun, OnUpdateStateFlags, ParseResponsePayload, ParseResponsePayloadLog, Reset
        MC_ReadActualForce/
          Structures/
            data type ReadActualForceOutCmd
            data type ReadActualForceParCmd
            data type ReadActualForceRecvData
            data type ReadActualForceSendData
          function block MC_ReadActualForceFB [ST]: CheckAddParameter, CheckFunctionSupported, CheckParameterChanged, CheckParameterValid, CreateCommandPayload, CreateCommandPayloadLog, FB_init, OnApplyOutCmd, OnExecRun, OnUpdateStateFlags, ParseResponsePayload, ParseResponsePayloadLog, Reset
      General/
        MC_CreateServerLog/
          Structures/
            data type CreateServerLogOutCmd
            data type CreateServerLogParCmd
            data type CreateServerLogRecvData
            data type CreateServerLogSendData
          function block MC_CreateServerLogFB [ST]: CheckAddParameter, CheckFunctionSupported, CheckParameterChanged, CheckParameterValid, CreateCommandPayload, CreateCommandPayloadLog, FB_init, OnApplyOutCmd, OnExecRun, OnUpdateStateFlags, ParseResponsePayload, ParseResponsePayloadLog, Reset
        MC_CreateServerLog_ToDo/
          function block MC_CreateServerLog_ToDo [ST]: FB_init
        MC_EnableRobot/
          Structures/
            data type EnableRobotOutCmd
            data type EnableRobotParCmd
            data type EnableRobotRecvData
            data type EnableRobotSendData
          function block MC_EnableRobotFB [ST]: CheckAddParameter, CheckFunctionSupported, CheckParameterChanged, CheckParameterValid, CheckSynchronizationValid, CreateCommandPayload, CreateCommandPayloadLog, FB_init, OnExecCancel, OnExecErrorClear, OnExecRun, OnUpdateStateFlags, ParseResponsePayload, ParseResponsePayloadLog, Reset
        MC_GroupReset/
          Structures/
            data type GroupResetOutCmd
            data type GroupResetParCmd
            data type GroupResetRecvData
            data type GroupResetSendData
          function block MC_GroupResetFB [ST]: CheckAddParameter, CheckFunctionSupported, CheckParameterChanged, CreateCommandPayload, CreateCommandPayloadLog, FB_init, OnExecRun, OnUpdateStateFlags, ParseResponsePayload, ParseResponsePayloadLog, Reset
        MC_ReadServerLog/
          Structures/
            data type ReadServerLogOutCmd
            data type ReadServerLogParCmd
            data type ReadServerLogRecvData
            data type ReadServerLogSendData
          function block MC_ReadServerLogFB [ST]: CheckAddParameter, CheckFunctionSupported, CheckParameterChanged, CheckParameterValid, CreateCommandPayload, CreateCommandPayloadLog, FB_init, OnApplyOutCmd, OnExecRun, OnUpdateStateFlags, ParseResponsePayload, ParseResponsePayloadLog, Reset, StoreLogContent
        MC_ReadServerLog_ToDo/
          function block MC_ReadServerLog [ST]: FB_init
        MC_RestartController/
          Structures/
            data type RestartControllerOutCmd
            data type RestartControllerParCmd
            data type RestartControllerRecvData
            data type RestartControllerSendData
          function block MC_RestartControllerFB [ST]: CheckAddParameter, CheckFunctionSupported, CheckParameterChanged, CreateCommandPayload, CreateCommandPayloadLog, FB_init, OnApplyOutCmd, OnExecRun, OnUpdateStateFlags, ParseResponsePayload, ParseResponsePayloadLog, Reset
        MC_RobotTask/
          Structures/
            ParCfg/
              Com/
                data type RobotTaskParCfgCom
              Plc/
                data type RobotTaskParCfgPlc
                data type RobotTaskParCfgPlcParameter
              Rob/
                data type RobotTaskParCfgRob
                data type RobotTaskParCfgRobParameter
              data type RobotTaskParCfg
          function block MC_RobotTaskFB [ST]: AxesGroupFromTelegram, AxesGroupFromTelegramCyclic, AxesGroupFromTelegramCyclicOptional, AxesGroupToTelegram, AxesGroupToTelegramCyclic, AxesGroupToTelegramCyclicOptional, AxesGroupToTelegramFooter, AxesGroupToTelegramHeader, AxesGroupToTelegramLogging, AxesGroupToTelegramSequence, CalculateCyclicDataLength, CalculateSequencePayloadMax, CalculateSequencePayloadStartAdr, CalculateTelegramLengthPlcToRob, CheckAssignmentValid, CheckParameterChanged, CheckParameterValid, CreateSendPayload, CreateSendPayloadCyclic, CreateSendPayloadCyclicOptional, CreateSendPayloadFooter, CreateSendPayloadHeader, CreateSendPayloadLogging, CreateSendPayloadSequence, FB_init, HandleAliveBit, HandleAxesGroup, HandleAxesGroupAcyclic, HandleAxesGroupCyclic, HandleAxesGroupCyclicOptional, HandleAxesGroupMessageLog, HandleAxesGroupParameter, HandleAxesGroupState, HandleAxesGroupSystemData, HandleInvalidFrames, HandleLifeSign, HandleLogMessagesAck, HandleSeqAck, HandleSync, HandleSyncFrameData, HandleSyncLoadData, HandleSyncRobotDefaultDynamics, HandleSyncRobotReferenceDynamics, HandleSyncRobotSWLimits, HandleSyncToolData, HandleSyncWorkArea, HandleTelegramStateCtrl, HandleUserData, HasError, HasInfo, HasWarning, OnCall, OnExecRun, ParseRecvPayload, ParseRecvPayloadCyclic, ParseRecvPayloadCyclicOptional, ParseRecvPayloadFooter, ParseRecvPayloadHeader, ParseRecvPayloadLogging, ParseRecvPayloadSequence, Reset, SetError, SetInfo, SetWarning, SyncModesValid
        MC_SetOperationMode/
          Structures/
            data type SetOperationModeOutCmd
            data type SetOperationModeParCmd
            data type SetOperationModeRecvData
            data type SetOperationModeSendData
          function block MC_SetOperationModeFB [ST]: CheckAddParameter, CheckFunctionSupported, CheckParameterChanged, CheckParameterValid, CreateCommandPayload, CreateCommandPayloadLog, FB_init, OnExecRun, OnUpdateStateFlags, ParseResponsePayload, ParseResponsePayloadLog, Reset
        MC_SetSequence/
          Structures/
            data type SetSequenceOutCmd
            data type SetSequenceParCmd
            data type SetSequenceRecvData
            data type SetSequenceSendData
          function block MC_SetSequenceFB [ST]: CheckAddParameter, CheckFunctionSupported, CheckParameterChanged, CheckParameterValid, CreateCommandPayload, CreateCommandPayloadLog, FB_init, OnExecRun, OnUpdateStateFlags, ParseResponsePayload, ParseResponsePayloadLog, Reset
        MC_SwitchLanguage/
          Structures/
            data type SwitchLanguageOutCmd
            data type SwitchLanguageParCmd
            data type SwitchLanguageRecvData
            data type SwitchLanguageSendData
          function block MC_SwitchLanguageFB [ST]: CheckAddParameter, CheckFunctionSupported, CheckParameterChanged, CheckParameterValid, CreateCommandPayload, CreateCommandPayloadLog, FB_init, OnApplyOutCmd, OnExecRun, OnUpdateStateFlags, ParseResponsePayload, ParseResponsePayloadLog, Reset
        MC_UserLogin/
          Structures/
            data type UserLoginOutCmd
            data type UserLoginParCmd
            data type UserLoginRecvData
            data type UserLoginSendData
          function block MC_UserLoginFB [ST]: CheckAddParameter, CheckFunctionSupported, CheckParameterChanged, CheckParameterValid, CreateCommandPayload, CreateCommandPayloadLog, FB_init, OnExecRun, OnUpdateStateFlags, ParseResponsePayload, ParseResponsePayloadLog, Reset
      Read/
        MC_ReadActualPosition/
          Structures/
            data type ReadActualPositionOutCmd
            data type ReadActualPositionParCmd
            data type ReadActualPositionRecvData
            data type ReadActualPositionSendData
          function block MC_ReadActualPositionFB [ST]: CheckAddParameter, CheckFunctionSupported, CheckParameterChanged, CheckParameterValid, CreateCommandPayload, CreateCommandPayloadLog, FB_init, OnApplyOutCmd, OnExecRun, OnUpdateStateFlags, ParseResponsePayload, ParseResponsePayloadLog, Reset
        MC_ReadActualPositionCyclic/
          Structures/
            data type ReadActualPositionCyclicOutCmd
            data type ReadActualPositionCyclicParCmd
          function block MC_ReadActualPositionCyclicFB [ST]: CheckFunctionSupported, CheckParameterChanged, CheckParameterValid, CreateCommandParameterLog, FB_init, OnCall, OnExecErrorClear, OnExecRun, Reset
        MC_ReadActualTCPVelocity/
          Structures/
            data type ReadActualTCPVelocityOutCmd
            data type ReadActualTCPVelocityParCmd
            data type ReadActualTCPVelocityRecvData
            data type ReadActualTCPVelocitySendData
          function block MC_ReadActualTCPVelocityFB [ST]: CheckAddParameter, CheckFunctionSupported, CheckParameterChanged, CheckParameterValid, CreateCommandPayload, CreateCommandPayloadLog, FB_init, OnApplyOutCmd, OnExecRun, OnUpdateStateFlags, ParseResponsePayload, ParseResponsePayloadLog, Reset
        MC_ReadAnalogInput/
          Structures/
            data type ReadAnalogInputOutCmd
            data type ReadAnalogInputParCmd
            data type ReadAnalogInputRecvData
            data type ReadAnalogInputSendData
          function block MC_ReadAnalogInputFB [ST]: CheckAddParameter, CheckFunctionSupported, CheckParameterChanged, CheckParameterValid, CreateCommandPayload, CreateCommandPayloadLog, FB_init, OnApplyOutCmd, OnExecRun, OnUpdateStateFlags, ParseResponsePayload, ParseResponsePayloadLog, Reset
        MC_ReadAnalogOutput/
          Structures/
            data type ReadAnalogOutputOutCmd
            data type ReadAnalogOutputParCmd
            data type ReadAnalogOutputRecvData
            data type ReadAnalogOutputSendData
          function block MC_ReadAnalogOutputFB [ST]: CheckAddParameter, CheckFunctionSupported, CheckParameterChanged, CheckParameterValid, CreateCommandPayload, CreateCommandPayloadLog, FB_init, OnApplyOutCmd, OnExecRun, OnUpdateStateFlags, ParseResponsePayload, ParseResponsePayloadLog, Reset
        MC_ReadDHParameter/
          Structures/
            data type ReadDHParameterOutCmd
            data type ReadDHParameterParCmd
            data type ReadDHParameterRecvData
            data type ReadDHParameterSendData
          function block MC_ReadDHParameterFB [ST]: CheckAddParameter, CheckFunctionSupported, CheckParameterChanged, CheckParameterValid, CreateCommandPayload, CreateCommandPayloadLog, FB_init, OnApplyOutCmd, OnExecRun, OnUpdateStateFlags, ParseResponsePayload, ParseResponsePayloadLog, Reset
        MC_ReadDigitalInputs/
          Structures/
            data type ReadDigitalInputsOutCmd
            data type ReadDigitalInputsParCmd
            data type ReadDigitalInputsRecvData
            data type ReadDigitalInputsSendData
          function block MC_ReadDigitalInputsFB [ST]: CheckAddParameter, CheckFunctionSupported, CheckParameterChanged, CheckParameterValid, CreateCommandPayload, CreateCommandPayloadLog, FB_init, OnApplyOutCmd, OnExecRun, OnUpdateStateFlags, ParseResponsePayload, ParseResponsePayloadLog, Reset
        MC_ReadDigitalOutputs/
          Structures/
            data type ReadDigitalOutputsOutCmd
            data type ReadDigitalOutputsParCmd
            data type ReadDigitalOutputsRecvData
            data type ReadDigitalOutputsSendData
          function block MC_ReadDigitalOutputsFB [ST]: CheckAddParameter, CheckFunctionSupported, CheckParameterChanged, CheckParameterValid, CreateCommandPayload, CreateCommandPayloadLog, FB_init, OnApplyOutCmd, OnExecRun, OnUpdateStateFlags, ParseResponsePayload, ParseResponsePayloadLog, Reset
        MC_ReadFrameData/
          Structures/
            data type ReadFrameDataOutCmd
            data type ReadFrameDataParCmd
            data type ReadFrameDataRecvData
            data type ReadFrameDataSendData
          function block MC_ReadFrameDataFB [ST]: CheckAddParameter, CheckFunctionSupported, CheckParameterChanged, CheckParameterValid, CreateCommandPayload, CreateCommandPayloadLog, FB_init, OnApplyOutCmd, OnExecRun, OnUpdateStateFlags, ParseResponsePayload, ParseResponsePayloadLog, Reset
        MC_ReadIntegers/
          Structures/
            data type ReadIntegersOutCmd
            data type ReadIntegersParCmd
            data type ReadIntegersRecvData
            data type ReadIntegersSendData
          function block MC_ReadIntegersFB [ST]: CheckAddParameter, CheckFunctionSupported, CheckParameterChanged, CheckParameterValid, CreateCommandPayload, CreateCommandPayloadLog, FB_init, OnApplyOutCmd, OnExecRun, OnUpdateStateFlags, ParseResponsePayload, ParseResponsePayloadLog, Reset
        MC_ReadLoadData/
          Structures/
            data type ReadLoadDataOutCmd
            data type ReadLoadDataParCmd
            data type ReadLoadDataRecvData
            data type ReadLoadDataSendData
          function block MC_ReadLoadDataFB [ST]: CheckAddParameter, CheckFunctionSupported, CheckParameterChanged, CheckParameterValid, CreateCommandPayload, CreateCommandPayloadLog, FB_init, OnApplyOutCmd, OnExecRun, OnUpdateStateFlags, ParseResponsePayload, ParseResponsePayloadLog, Reset
        MC_ReadMessages/
          Structures/
            data type ReadMessagesOutCmd
            data type ReadMessagesParCmd
            data type ReadMessagesRecvData
            data type ReadMessagesSendData
          function block MC_ReadMessagesFB [ST]: CheckAddParameter, CheckFunctionSupported, CheckParameterChanged, CheckParameterValid, CreateCommandPayload, CreateCommandPayloadLog, FB_init, OnApplyOutCmd, OnExecCancel, OnExecErrorClear, OnExecRun, OnUpdateStateFlags, ParseResponsePayload, ParseResponsePayloadLog, Reset
        MC_ReadReals/
          Structures/
            data type ReadRealsOutCmd
            data type ReadRealsParCmd
            data type ReadRealsRecvData
            data type ReadRealsSendData
          function block MC_ReadRealsFB [ST]: CheckAddParameter, CheckFunctionSupported, CheckParameterChanged, CheckParameterValid, CreateCommandPayload, CreateCommandPayloadLog, FB_init, OnApplyOutCmd, OnExecRun, OnUpdateStateFlags, ParseResponsePayload, ParseResponsePayloadLog, Reset
        MC_ReadRobotData/
          Structures/
            data type ReadRobotDataOutCmd
            data type ReadRobotDataParCmd
            data type ReadRobotDataRecvData
            data type ReadRobotDataSendData
          function block MC_ReadRobotDataFB [ST]: CheckAddParameter, CheckFunctionSupported, CheckParameterChanged, CreateCommandPayload, CreateCommandPayloadLog, FB_init, OnApplyOutCmd, OnExecRun, OnUpdateStateFlags, ParseResponsePayload, ParseResponsePayloadLog, Reset
        MC_ReadRobotDefaultDynamics/
          Structures/
            data type ReadRobotDefaultDynamicsOutCmd
            data type ReadRobotDefaultDynamicsParCmd
            data type ReadRobotDefaultDynamicsRecvData
            data type ReadRobotDefaultDynamicsSendData
          function block MC_ReadRobotDefaultDynamicsFB [ST]: CheckAddParameter, CheckFunctionSupported, CheckParameterChanged, CreateCommandPayload, CreateCommandPayloadLog, FB_init, OnApplyOutCmd, OnExecRun, OnUpdateStateFlags, ParseResponsePayload, ParseResponsePayloadLog, Reset
        MC_ReadRobotReferenceDynamics/
          Structures/
            data type ReadRobotReferenceDynamicsOutCmd
            data type ReadRobotReferenceDynamicsParCmd
            data type ReadRobotReferenceDynamicsRecvData
            data type ReadRobotReferenceDynamicsSendData
          function block MC_ReadRobotReferenceDynamicsFB [ST]: CheckAddParameter, CheckFunctionSupported, CheckParameterChanged, CreateCommandPayload, CreateCommandPayloadLog, FB_init, OnApplyOutCmd, OnExecRun, OnUpdateStateFlags, ParseResponsePayload, ParseResponsePayloadLog, Reset
        MC_ReadRobotSWLimits/
          Structures/
            data type ReadRobotSWLimitsOutCmd
            data type ReadRobotSWLimitsParCmd
            data type ReadRobotSWLimitsRecvData
            data type ReadRobotSWLimitsSendData
          function block MC_ReadRobotSWLimitsFB [ST]: CheckAddParameter, CheckFunctionSupported, CheckParameterChanged, CreateCommandPayload, CreateCommandPayloadLog, FB_init, OnApplyOutCmd, OnExecRun, OnUpdateStateFlags, ParseResponsePayload, ParseResponsePayloadLog, Reset
        MC_ReadSystemVariable/
          Structures/
            data type ReadSystemVariableOutCmd
            data type ReadSystemVariableParCmd
            data type ReadSystemVariableRecvData
            data type ReadSystemVariableSendData
          function block MC_ReadSystemVariableFB [ST]: CheckAddParameter, CheckFunctionSupported, CheckParameterChanged, CheckParameterValid, CreateCommandPayload, CreateCommandPayloadLog, FB_init, OnApplyOutCmd, OnExecRun, OnUpdateStateFlags, ParseResponsePayload, ParseResponsePayloadLog, Reset
        MC_ReadToolData/
          Structures/
            data type ReadToolDataOutCmd
            data type ReadToolDataParCmd
            data type ReadToolDataRecvData
            data type ReadToolDataSendData
          function block MC_ReadToolDataFB [ST]: CheckAddParameter, CheckFunctionSupported, CheckParameterChanged, CheckParameterValid, CreateCommandPayload, CreateCommandPayloadLog, FB_init, OnApplyOutCmd, OnExecRun, OnUpdateStateFlags, ParseResponsePayload, ParseResponsePayloadLog, Reset
      SearchHardstop/
        MC_SearchHardStop/
          Structures/
            data type SearchHardStopOutCmd
            data type SearchHardStopParCmd
            data type SearchHardStopRecvData
            data type SearchHardStopSendData
          function block MC_SearchHardStopFB [ST]: CheckAddParameter, CheckFunctionSupported, CheckParameterChanged, CheckParameterValid, CreateCommandPayload, CreateCommandPayloadLog, FB_init, OnApplyOutCmd, OnExecRun, OnUpdateStateFlags, ParseResponsePayload, ParseResponsePayloadLog, Reset
        MC_SearchHardStopJ/
          Structures/
            data type SearchHardStopJOutCmd
            data type SearchHardStopJParCmd
            data type SearchHardStopJRecvData
            data type SearchHardStopJSendData
          function block MC_SearchHardStopJFB [ST]: CheckAddParameter, CheckFunctionSupported, CheckParameterChanged, CheckParameterValid, CreateCommandPayload, CreateCommandPayloadLog, FB_init, OnApplyOutCmd, OnExecRun, OnUpdateStateFlags, ParseResponsePayload, ParseResponsePayloadLog, Reset
      Spline/
        MC_CreateSpline/
          Structures/
            data type CreateSplineOutCmd
            data type CreateSplineParCmd
            data type CreateSplineRecvData
            data type CreateSplineSendData
          function block MC_CreateSplineFB [ST]: CheckAddParameter, CheckFunctionSupported, CheckParameterChanged, CheckParameterValid, CreateCommandPayload, CreateCommandPayloadLog, FB_init, OnExecRun, OnUpdateStateFlags, ParseResponsePayload, ParseResponsePayloadLog, Reset
        MC_DeleteSpline/
          Structures/
            data type DeleteSplineOutCmd
            data type DeleteSplineParCmd
            data type DeleteSplineRecvData
            data type DeleteSplineSendData
          function block MC_DeleteSplineFB [ST]: CheckAddParameter, CheckFunctionSupported, CheckParameterChanged, CheckParameterValid, CreateCommandPayload, CreateCommandPayloadLog, FB_init, OnExecRun, OnUpdateStateFlags, ParseResponsePayload, ParseResponsePayloadLog, Reset
        MC_DynamicSpline/
          Structures/
            data type DynamicSplineOutCmd
            data type DynamicSplineParCmd
            data type DynamicSplineRecvData
            data type DynamicSplineSendData
          function block MC_DynamicSplineFB [ST]: CheckAddParameter, CheckFunctionSupported, CheckParameterChanged, CheckParameterValid, CreateCommandPayload, CreateCommandPayloadLog, FB_init, OnApplyOutCmd, OnExecCancel, OnExecErrorClear, OnExecRun, OnUpdateStateFlags, ParseResponsePayload, ParseResponsePayloadLog, Reset
        MC_MoveSpline/
          Structures/
            data type MoveSplineOutCmd
            data type MoveSplineParCmd
            data type MoveSplineRecvData
            data type MoveSplineSendData
          function block MC_MoveSplineFB [ST]: CheckAddParameter, CheckFunctionSupported, CheckParameterChanged, CheckParameterValid, CreateCommandPayload, CreateCommandPayloadLog, FB_init, OnApplyOutCmd, OnExecRun, OnUpdateStateFlags, ParseResponsePayload, ParseResponsePayloadLog, Reset
      SuperImposing/
        MC_MoveSuperImposed/
          Structures/
            data type MoveSuperImposedOutCmd
            data type MoveSuperImposedParCmd
            data type MoveSuperImposedRecvData
            data type MoveSuperImposedSendData
          function block MC_MoveSuperImposedFB [ST]: CheckAddParameter, CheckFunctionSupported, CheckParameterChanged, CheckParameterValid, CreateCommandPayload, CreateCommandPayloadLog, FB_init, OnApplyOutCmd, OnExecRun, OnUpdateStateFlags, ParseResponsePayload, ParseResponsePayloadLog, Reset
        MC_MoveSuperImposedDynamic/
          Structures/
            data type MoveSuperImposedDynamicOutCmd
            data type MoveSuperImposedDynamicParCmd
            data type MoveSuperImposedDynamicRecvData
            data type MoveSuperImposedDynamicSendData
          function block MC_MoveSuperImposedDynamicFB [ST]: CheckAddParameter, CheckFunctionSupported, CheckParameterChanged, CheckParameterValid, CreateCommandPayload, CreateCommandPayloadLog, FB_init, OnApplyOutCmd, OnExecRun, OnUpdateStateFlags, ParseResponsePayload, ParseResponsePayloadLog, Reset
      Trigger/
        MC_ReactAtTrigger/
          Structures/
            data type ReactAtTriggerOutCmd
            data type ReactAtTriggerParCmd
            data type ReactAtTriggerRecvData
            data type ReactAtTriggerSendData
          function block MC_ReactAtTriggerFB [ST]: CheckAddParameter, CheckFunctionSupported, CheckParameterChanged, CheckParameterValid, CreateCommandPayload, CreateCommandPayloadLog, FB_init, OnApplyOutCmd, OnExecRun, OnUpdateStateFlags, ParseResponsePayload, ParseResponsePayloadLog, Reset
        MC_SetTriggerError/
          Structures/
            data type SetTriggerErrorOutCmd
            data type SetTriggerErrorParCmd
            data type SetTriggerErrorRecvData
            data type SetTriggerErrorSendData
          function block MC_SetTriggerErrorFB [ST]: CheckAddParameter, CheckFunctionSupported, CheckParameterChanged, CheckParameterValid, CreateCommandPayload, CreateCommandPayloadLog, FB_init, OnApplyOutCmd, OnExecRun, OnUpdateStateFlags, ParseResponsePayload, ParseResponsePayloadLog, Reset
        MC_SetTriggerLimit/
          Structures/
            data type SetTriggerLimitOutCmd
            data type SetTriggerLimitParCmd
            data type SetTriggerLimitRecvData
            data type SetTriggerLimitSendData
          function block MC_SetTriggerLimitFB [ST]: CheckAddParameter, CheckFunctionSupported, CheckParameterChanged, CheckParameterValid, CreateCommandPayload, CreateCommandPayloadLog, FB_init, OnApplyOutCmd, OnExecRun, OnUpdateStateFlags, ParseResponsePayload, ParseResponsePayloadLog, Reset
        MC_SetTriggerMotion/
          Structures/
            data type SetTriggerMotionOutCmd
            data type SetTriggerMotionParCmd
            data type SetTriggerMotionRecvData
            data type SetTriggerMotionSendData
          function block MC_SetTriggerMotionFB [ST]: CheckAddParameter, CheckFunctionSupported, CheckParameterChanged, CheckParameterValid, CreateCommandPayload, CreateCommandPayloadLog, FB_init, OnApplyOutCmd, OnExecRun, OnUpdateStateFlags, ParseResponsePayload, ParseResponsePayloadLog, Reset
        MC_SetTriggerRegister/
          Structures/
            data type SetTriggerRegisterOutCmd
            data type SetTriggerRegisterParCmd
            data type SetTriggerRegisterRecvData
            data type SetTriggerRegisterSendData
          function block MC_SetTriggerRegisterFB [ST]: CheckAddParameter, CheckFunctionSupported, CheckParameterChanged, CheckParameterValid, CreateCommandPayload, CreateCommandPayloadLog, FB_init, OnApplyOutCmd, OnExecRun, OnUpdateStateFlags, ParseResponsePayload, ParseResponsePayloadLog, Reset
        MC_SetTriggerUser/
          Structures/
            data type SetTriggerUserOutCmd
            data type SetTriggerUserParCmd
            data type SetTriggerUserRecvData
            data type SetTriggerUserSendData
          function block MC_SetTriggerUserFB [ST]: CheckAddParameter, CheckFunctionSupported, CheckParameterChanged, CheckParameterValid, CreateCommandPayload, CreateCommandPayloadLog, FB_init, OnApplyOutCmd, OnExecRun, OnUpdateStateFlags, ParseResponsePayload, ParseResponsePayloadLog, Reset
        MC_WaitForTrigger/
          Structures/
            data type WaitForTriggerOutCmd
            data type WaitForTriggerParCmd
            data type WaitForTriggerRecvData
            data type WaitForTriggerSendData
          function block MC_WaitForTriggerFB [ST]: CheckAddParameter, CheckFunctionSupported, CheckParameterChanged, CheckParameterValid, CreateCommandPayload, CreateCommandPayloadLog, FB_init, OnApplyOutCmd, OnExecRun, OnUpdateStateFlags, ParseResponsePayload, ParseResponsePayloadLog, Reset
        MC_WaitTime/
          Structures/
            data type WaitTimeOutCmd
            data type WaitTimeParCmd
            data type WaitTimeRecvData
            data type WaitTimeSendData
          function block MC_WaitTimeFB [ST]: CheckAddParameter, CheckFunctionSupported, CheckParameterChanged, CheckParameterValid, CreateCommandPayload, CreateCommandPayloadLog, FB_init, OnApplyOutCmd, OnExecRun, OnUpdateStateFlags, ParseResponsePayload, ParseResponsePayloadLog, Reset
      WorkAreas/
        MC_ActivateWorkArea/
          Structures/
            data type ActivateWorkAreaOutCmd
            data type ActivateWorkAreaParCmd
            data type ActivateWorkAreaRecvData
            data type ActivateWorkAreaSendData
          function block MC_ActivateWorkAreaFB [ST]: CheckAddParameter, CheckFunctionSupported, CheckParameterChanged, CheckParameterValid, CreateCommandPayload, CreateCommandPayloadLog, FB_init, OnExecRun, OnUpdateStateFlags, ParseResponsePayload, ParseResponsePayloadLog, Reset
        MC_MonitorWorkArea/
          Structures/
            data type MonitorWorkAreaOutCmd
            data type MonitorWorkAreaParCmd
            data type MonitorWorkAreaRecvData
            data type MonitorWorkAreaSendData
          function block MC_MonitorWorkAreaFB [ST]: CheckAddParameter, CheckFunctionSupported, CheckParameterChanged, CheckParameterValid, CreateCommandPayload, CreateCommandPayloadLog, FB_init, OnApplyOutCmd, OnExecRun, OnUpdateStateFlags, ParseResponsePayload, ParseResponsePayloadLog, Reset
        MC_ReadWorkArea/
          Structures/
            data type ReadWorkAreaOutCmd
            data type ReadWorkAreaParCmd
            data type ReadWorkAreaRecvData
            data type ReadWorkAreaSendData
          function block MC_ReadWorkAreaFB [ST]: CheckAddParameter, CheckFunctionSupported, CheckParameterChanged, CheckParameterValid, CreateCommandPayload, CreateCommandPayloadLog, FB_init, OnApplyOutCmd, OnExecRun, OnUpdateStateFlags, ParseResponsePayload, ParseResponsePayloadLog, Reset
        MC_WriteWorkArea/
          Structures/
            data type WriteWorkAreaOutCmd
            data type WriteWorkAreaParCmd
            data type WriteWorkAreaRecvData
            data type WriteWorkAreaSendData
          function block MC_WriteWorkAreaFB [ST]: CheckAddParameter, CheckFunctionSupported, CheckParameterChanged, CheckParameterValid, CreateCommandPayload, CreateCommandPayloadLog, FB_init, OnExecRun, OnUpdateStateFlags, ParseResponsePayload, ParseResponsePayloadLog, Reset
      Write/
        MC_WriteAnalogOutput/
          Structures/
            data type WriteAnalogOutputOutCmd
            data type WriteAnalogOutputParCmd
            data type WriteAnalogOutputRecvData
            data type WriteAnalogOutputSendData
          function block MC_WriteAnalogOutputFB [ST]: CheckAddParameter, CheckFunctionSupported, CheckParameterChanged, CheckParameterValid, CreateCommandPayload, CreateCommandPayloadLog, FB_init, OnApplyOutCmd, OnExecRun, OnUpdateStateFlags, ParseResponsePayload, ParseResponsePayloadLog, Reset
        MC_WriteDigitalOutputs/
          Structures/
            data type WriteDigitalOutputsOutCmd
            data type WriteDigitalOutputsParCmd
            data type WriteDigitalOutputsRecvData
            data type WriteDigitalOutputsSendData
          function block MC_WriteDigitalOutputsFB [ST]: CheckAddParameter, CheckFunctionSupported, CheckParameterChanged, CheckParameterValid, CreateCommandPayload, CreateCommandPayloadLog, FB_init, OnApplyOutCmd, OnExecRun, OnUpdateStateFlags, ParseResponsePayload, ParseResponsePayloadLog, Reset
        MC_WriteFrameData/
          Structures/
            data type WriteFrameDataOutCmd
            data type WriteFrameDataParCmd
            data type WriteFrameDataRecvData
            data type WriteFrameDataSendData
          function block MC_WriteFrameDataFB [ST]: CheckAddParameter, CheckFunctionSupported, CheckParameterChanged, CheckParameterValid, CreateCommandPayload, CreateCommandPayloadLog, FB_init, OnExecRun, OnUpdateStateFlags, ParseResponsePayload, ParseResponsePayloadLog, Reset
        MC_WriteIntegers/
          Structures/
            data type WriteIntegersOutCmd
            data type WriteIntegersParCmd
            data type WriteIntegersRecvData
            data type WriteIntegersSendData
          function block MC_WriteIntegersFB [ST]: CheckAddParameter, CheckFunctionSupported, CheckParameterChanged, CheckParameterValid, CreateCommandPayload, CreateCommandPayloadLog, FB_init, OnApplyOutCmd, OnExecRun, OnUpdateStateFlags, ParseResponsePayload, ParseResponsePayloadLog, Reset
        MC_WriteLoadData/
          Structures/
            data type WriteLoadDataOutCmd
            data type WriteLoadDataParCmd
            data type WriteLoadDataRecvData
            data type WriteLoadDataSendData
          function block MC_WriteLoadDataFB [ST]: CheckAddParameter, CheckFunctionSupported, CheckParameterChanged, CheckParameterValid, CreateCommandPayload, CreateCommandPayloadLog, FB_init, OnExecRun, OnUpdateStateFlags, ParseResponsePayload, ParseResponsePayloadLog, Reset
        MC_WriteReals/
          Structures/
            data type WriteRealsOutCmd
            data type WriteRealsParCmd
            data type WriteRealsRecvData
            data type WriteRealsSendData
          function block MC_WriteRealsFB [ST]: CheckAddParameter, CheckFunctionSupported, CheckParameterChanged, CheckParameterValid, CreateCommandPayload, CreateCommandPayloadLog, FB_init, OnApplyOutCmd, OnExecRun, OnUpdateStateFlags, ParseResponsePayload, ParseResponsePayloadLog, Reset
        MC_WriteRobotDefaultDynamics/
          Structures/
            data type WriteRobotDefaultDynamicsOutCmd
            data type WriteRobotDefaultDynamicsParCmd
            data type WriteRobotDefaultDynamicsRecvData
            data type WriteRobotDefaultDynamicsSendData
          function block MC_WriteRobotDefaultDynamicsFB [ST]: CheckAddParameter, CheckFunctionSupported, CheckParameterChanged, CheckParameterValid, CreateCommandPayload, CreateCommandPayloadLog, FB_init, OnApplyOutCmd, OnExecRun, OnUpdateStateFlags, ParseResponsePayload, ParseResponsePayloadLog, Reset
        MC_WriteRobotReferenceDynamics/
          Structures/
            data type WriteRobotReferenceDynamicsOutCmd
            data type WriteRobotReferenceDynamicsParCmd
            data type WriteRobotReferenceDynamicsRecvData
            data type WriteRobotReferenceDynamicsSendData
          function block MC_WriteRobotReferenceDynamicsFB [ST]: CheckAddParameter, CheckFunctionSupported, CheckParameterChanged, CheckParameterValid, CreateCommandPayload, CreateCommandPayloadLog, FB_init, OnApplyOutCmd, OnExecRun, OnUpdateStateFlags, ParseResponsePayload, ParseResponsePayloadLog, Reset
        MC_WriteRobotSWLimits/
          Structures/
            data type WriteRobotSWLimitsOutCmd
            data type WriteRobotSWLimitsParCmd
            data type WriteRobotSWLimitsRecvData
            data type WriteRobotSWLimitsSendData
          function block MC_WriteRobotSWLimitsFB [ST]: CheckAddParameter, CheckFunctionSupported, CheckParameterChanged, CheckParameterValid, CreateCommandPayload, CreateCommandPayloadLog, FB_init, OnApplyOutCmd, OnExecRun, OnUpdateStateFlags, ParseResponsePayload, ParseResponsePayloadLog, Reset
        MC_WriteSystemVariable/
          Structures/
            data type WriteSystemVariableOutCmd
            data type WriteSystemVariableParCmd
            data type WriteSystemVariableRecvData
            data type WriteSystemVariableSendData
          function block MC_WriteSystemVariableFB [ST]: CheckAddParameter, CheckFunctionSupported, CheckParameterChanged, CheckParameterValid, CreateCommandPayload, CreateCommandPayloadLog, FB_init, OnApplyOutCmd, OnExecRun, OnUpdateStateFlags, ParseResponsePayload, ParseResponsePayloadLog, Reset
        MC_WriteToolData/
          Structures/
            data type WriteToolDataOutCmd
            data type WriteToolDataParCmd
            data type WriteToolDataRecvData
            data type WriteToolDataSendData
          function block MC_WriteToolDataFB [ST]: CheckAddParameter, CheckFunctionSupported, CheckParameterChanged, CheckParameterValid, CreateCommandPayload, CreateCommandPayloadLog, FB_init, OnExecRun, OnUpdateStateFlags, ParseResponsePayload, ParseResponsePayloadLog, Reset
    Structures/
      _internal/
        data type SplineDataSend
      AxesGroup/
        Acyclic/
          data type AxesGroupAcyclic
          data type AxesGroupAcyclicAcrEntry
          data type AxesGroupAcyclicAcrEntryCmdBuffer
          data type AxesGroupAcyclicAcrEntryRspBuffer
          data type AxesGroupAcyclicExecutionOrderList
        Cyclic/
          data type AxesGroupCyclic
          data type AxesGroupCyclicPlcToRob
          data type AxesGroupCyclicRobToPlc
        CyclicOptional/
          Internal/
            data type AxesGroupCyclicOptionalDataCartesianPosition
            data type AxesGroupCyclicOptionalDataCartesianPositionExt
            data type AxesGroupCyclicOptionalDataCurrent
            data type AxesGroupCyclicOptionalDataCurrentExt
            data type AxesGroupCyclicOptionalDataForce
            data type AxesGroupCyclicOptionalDataForceExt
            data type AxesGroupCyclicOptionalDataJointPosition
            data type AxesGroupCyclicOptionalDataJointPositionExt
            data type AxesGroupCyclicOptionalDataSubProgram
          data type AxesGroupCyclicOptionalData
          data type AxesGroupCyclicOptionalDataPlcToRob
          data type AxesGroupCyclicOptionalDataRobToPlc
        MessageLog/
          data type AxesGroupMessageLog
        Parameter/
          OptionalCyclic/
            data type AxesGroupParameterOptionalCyclic
            data type AxesGroupParameterOptionalCyclicPlcToRob
            data type AxesGroupParameterOptionalCyclicRobToPlc
          Plc/
            data type AxesGroupParameterPlc
            data type AxesGroupParameterPlcOptionalCyclic
            data type AxesGroupParameterPlcParameter
          Rob/
            data type AxesGroupParameterRob
            data type AxesGroupParameterRobOptionalCyclic
            data type AxesGroupParameterRobParameter
          data type AxesGroupParameter
        State/
          DataChanged/
            data type AxesGroupStateDataChanged
          Synchronizing/
            data type AxesGroupStateSynchronizing
          SyncState/
            data type AxesGroupStateSyncState
            data type AxesGroupStateSyncStateNo
            data type AxesGroupStateSyncStatePlc
            data type AxesGroupStateSyncStateRob
          data type AxesGroupState
        data type AxesGroup
      Axis/
        data type AxisExternalUnit
        data type AxisExternalUsed
        data type AxisJointUnit
        data type AxisJointUsed
      Cartesian/
        data type RobotCartesianForce
        data type RobotCartesianForceExt
        data type RobotCartesianForceShort
        data type RobotCartesianPosition
        data type RobotCartesianPositionBase
        data type RobotCartesianPositionExt
        data type RobotCartesianPositionShort
      Common/
        data type CmdHeader
        data type LogParameter
        data type RobotCoordinateSystemParameters
        data type RspHeader
      Data/
        Frame/
          data type Frame
          data type FrameData
        Load/
          data type Load
          data type LoadData
        Spline/
          data type SplineData
        SubProgram/
          data type RobotSubProgramData
        Tool/
          data type Tool
          data type ToolData
        User/
          data type UserData
        WorkArea/
          data type RobotWorkArea
          data type RobotWorkAreaData
          data type RobotWorkAreaDataLimitCartesian
          data type RobotWorkAreaDataLimitJoint
        data type CyclicStateData
      DatenAndTime/
        data type IEC_DATE
        data type IEC_TIME
        data type IEC_TIMESTAMP
        data type SystemTime
      Dynamics/
        data type DefaultDynamics
        data type ReferenceDynamics
        data type RobotDynamics
      Joint/
        data type RobotJointCurrent
        data type RobotJointCurrentExt
        data type RobotJointCurrentShort
        data type RobotJointPosition
        data type RobotJointPositionExt
        data type RobotJointPositionShort
      Miscellaneous/
        data type AlarmMessage
        data type ArmConfigParameter
        data type AuxOffset
        data type CoordinateSystem
        data type DataEnableSync
        data type DataInSync
        data type DHParameter
        data type ExecutionModeAllowed
        data type ExternalAxesFlags
        data type ForceStatus
        data type FragmentAction
        data type JogControl
        data type MeasuringInputResult
        data type ProcessingModeAllowed
        data type RaStatusWord
        data type RCSupportedFunctions
        data type RobotAxesFlags
        data type SWLimits
        data type SynchronizationModes
        data type SyncUserInteraction
        data type TrackingStatus
        data type TurnNumber
        data type VersionStruct
      Telegram/
        PlcToRob/
          Command/
            data type TelegramPlcToRobCommand
            data type TelegramPlcToRobCommandHeader
          Cyclic/
            data type TelegramPlcToRobCyclicData
          CyclicOptional/
            Internal/
              data type TelegramPlcToRobCyclicOptionalCartesianPosition
              data type TelegramPlcToRobCyclicOptionalCartesianPositionExt
              data type TelegramPlcToRobCyclicOptionalCurrent
              data type TelegramPlcToRobCyclicOptionalCurrentExt
              data type TelegramPlcToRobCyclicOptionalForce
              data type TelegramPlcToRobCyclicOptionalForceExt
              data type TelegramPlcToRobCyclicOptionalJointPosition
              data type TelegramPlcToRobCyclicOptionalJointPositionExt
              data type TelegramPlcToRobCyclicOptionalSubProgramData
            data type TelegramPlcToRobCyclicOptionalData
          Footer/
            data type TelegramPlcToRobFooter
          Fragment/
            data type TelegramPlcToRobFragment
            data type TelegramPlcToRobFragmentHeader
          Header/
            data type TelegramPlcToRobHeader
          Sequence/
            data type TelegramPlcToRobSequence
            data type TelegramPlcToRobSequenceHeader
          data type TelegramPlcToRob
        RobToPlc/
          Command/
            data type TelegramRobToPlcCommand
            data type TelegramRobToPlcCommandHeader
          CyclicOptional/
            Internal/
              data type TelegramRobToPlcCyclicOptionalCartesianPosition
              data type TelegramRobToPlcCyclicOptionalCartesianPositionExt
              data type TelegramRobToPlcCyclicOptionalCurrent
              data type TelegramRobToPlcCyclicOptionalCurrentExt
              data type TelegramRobToPlcCyclicOptionalForce
              data type TelegramRobToPlcCyclicOptionalForceExt
              data type TelegramRobToPlcCyclicOptionalJointPosition
              data type TelegramRobToPlcCyclicOptionalJointPositionExt
              data type TelegramRobToPlcCyclicOptionalSubProgramData
            data type TelegramRobToPlcCyclicOptionalData
          Footer/
            data type TelegramRobToPlcFooter
          Fragment/
            data type TelegramRobToPlcFragment
            data type TelegramRobToPlcFragmentHeader
          Header/
            data type TelegramRobToPlcHeader
          Sequence/
            data type TelegramRobToPlcSequence
            data type TelegramRobToPlcSequenceHeader
          data type TelegramRobToPlc
        data type Telegram
*)

// Library/Enumerations/ArmConfig/ArmConfigElbow
{attribute 'qualified_only'}
// {attribute 'to_string'} // bth3ho Fanuc
// ------------------------------------------------------------------------- 
//  SRCI Robot Library                                                
// ------------------------------------------------------------------------- 
//                                                                           
//  Object:      ArmConfigElbow                                       
//  Author:      Thorsten Brach                                                
//  Date:        2024-06-01
//
//  Description:                                              
//   
//                                                                           
//  Copyright: 
//    (C) 2024 Thorsten Brach. All rights reserved                                                                                                                                            
//             Licensed under the MIT License.
//                                                                           
//  Disclaimer:                                                                           
//    This project is provided without any guarantee and can be used for   
//    private and commercial purposes. Any use is at the user’s 
//    own risk and responsibility.
//
// -------------------------------------------------------------------------
TYPE ArmConfigElbow :
(
 /// Use config in position  
 USE_CONFIG := 0,
 /// Do not change config with this movement. (default)
 SAME := 1,
 /// Configuration in position is not used but the Robot is free to change config
 FREE := 2,
 /// Set elbow configuration in position to Down
 DOWN := 3,
 /// Set elbow configuration in position to up
 UP := 4
);
END_TYPE

// Library/Enumerations/ArmConfig/ArmConfigShoulder
{attribute 'qualified_only'}
// {attribute 'to_string'} // bth3ho Fanuc
// ------------------------------------------------------------------------- 
//  SRCI Robot Library                                                
// ------------------------------------------------------------------------- 
//                                                                           
//  Object:      ArmConfigShoulder                                       
//  Author:      Thorsten Brach                                                
//  Date:        2024-06-01
//
//  Description:                                              
//   
//                                                                           
//  Copyright: 
//    (C) 2024 Thorsten Brach. All rights reserved                                                                                                                                            
//             Licensed under the MIT License.
//                                                                           
//  Disclaimer:                                                                           
//    This project is provided without any guarantee and can be used for   
//    private and commercial purposes. Any use is at the user’s 
//    own risk and responsibility.
//
// -------------------------------------------------------------------------
TYPE ArmConfigShoulder :
(
 /// Use config in position  
 USE_CONFIG := 0,
 /// Do not change config with this movement. (default)
 SAME := 1,
 /// Configuration in position is not used but the Robot is free to change config
 FREE := 2,
 /// Set shoulder configuration in position to Back
 BACK := 3,
 /// Set shoulder configuration in position to Front
 FRONT := 4
);
END_TYPE

// Library/Enumerations/ArmConfig/ArmConfigWrist
{attribute 'qualified_only'}
// {attribute 'to_string'} // bth3ho Fanuc
// ------------------------------------------------------------------------- 
//  SRCI Robot Library                                                
// ------------------------------------------------------------------------- 
//                                                                           
//  Object:      ArmConfigWrist                                       
//  Author:      Thorsten Brach                                                
//  Date:        2024-06-01
//
//  Description:                                              
//   
//                                                                           
//  Copyright: 
//    (C) 2024 Thorsten Brach. All rights reserved                                                                                                                                            
//             Licensed under the MIT License.
//                                                                           
//  Disclaimer:                                                                           
//    This project is provided without any guarantee and can be used for   
//    private and commercial purposes. Any use is at the user’s 
//    own risk and responsibility.
//
// -------------------------------------------------------------------------
TYPE ArmConfigWrist :
(
 /// Use config in position  
 USE_CONFIG := 0,
 /// Do not change config with this movement. (default)
 SAME := 1,
 /// Configuration in position is not used but the Robot is free to change config
 FREE := 2,
 /// Set wrist configuration in position to Flip
 FLIP := 3,
 /// Set wrist configuration in position to Non-Flip
 NON_FLIP := 4
);
END_TYPE

// Library/Enumerations/Events/RobotLibraryErrorIdEnum
{attribute 'qualified_only'}
{attribute 'to_string'}
// ------------------------------------------------------------------------- 
//  SRCI Robot Library                                                
// ------------------------------------------------------------------------- 
//                                                                           
//  Object:      RobotLibraryErrorIdEnum                                       
//  Author:      Thorsten Brach                                                
//  Date:        2024-06-01
//
//  Description:                                              
//   
//                                                                           
//  Copyright: 
//    (C) 2024 Thorsten Brach. All rights reserved                                                                                                                                            
//             Licensed under the MIT License.
//                                                                           
//  Disclaimer:                                                                           
//    This project is provided without any guarantee and can be used for   
//    private and commercial purposes. Any use is at the user’s 
//    own risk and responsibility.
//
// -------------------------------------------------------------------------
TYPE RobotLibraryErrorIdEnum :
(
  NO_ERROR := 0,

  {warning 'ToDo: This is an internal error ID, which is not defined in SRCI specification'}
  /// START
  
  /// Program fault : Invalid step
  ERR_INVALID_STEP             := 1,
  /// Program fault : Invalid library parameter
  ERR_INVALID_LIBRARY_PARA     := 2,
  /// Program fault : Invalid axes groups ID
  ERR_INVALID_AXES_GROUP_ID    := 3,

  /// Function is not supported
  ERR_FUNCTION_NOT_SUPPORTED   := 5,
  /// Program fault : Timeout during command execution 
  ERR_TIMEOUT_CMD              := 6,
  /// Parameter fault : Invalid command parameter SyncReaction
  ERR_INVALID_PAR_CMD_SYNC_REACTION  := 7,
  /// Invalid command parameter - see log file for details (LogLevel Error)
  ERR_INVALID_PAR_CMD := 8,             
  /// Synchronisation state prohibits command execution
  ERR_SYNC_STATE_PROHIBITS_COMMAND := 9,
  // ST-FIX F130: ERR_SYNC_MODE_INVALID (10) removed - an invalid SyncMode is only a warning (WARN_*_SYNC_MODE_INVALID)
  /// Client Invalid parameter value - LoadNo not
  /// available on RC
  /// Commands using the parameter "LoadNo"
  ERR_LOADNO_UNAVAILABLE  := 11,   
  /// Client Invalid parameter value - WorkAreaNo outside of
  /// the allowed range -1..254
  /// Commands using the parameter "WorkAreaNo"
  ERR_WORKAREANO_RANGE  := 12,
  /// Client Invalid parameter value - LoadNo not
  /// available on RC
  /// Commands using the parameter "LoadNo"
  ERR_WORKAREANO_UNAVAILABLE  := 13,   
  /// Client Specified TriggerMode not allowed
  /// Commands using the parameter "TriggerMode"
  ERR_TRIGGERMODE_NOT_ALLOWED := 14, 
  /// Client Specified Frame calculation mode not valid
  /// Commands using the parameter "FrameCalculationMode"
  ERR_FRAMECALCULATIONMODE_INVALID := 15,

  /// RC tool count higher than PLC tool count -> Synchronization not possible 
  ERR_SYNC_TOOL_COUNT_RC_HIGHER_THAN_PLC := 16,
  /// RC load count higher than PLC load count -> Synchronization not possible 
  ERR_SYNC_LOAD_COUNT_RC_HIGHER_THAN_PLC := 17,
  /// RC frame count higher than PLC frame count -> Synchronization not possible 
  ERR_SYNC_FRAME_COUNT_RC_HIGHER_THAN_PLC := 18,
  /// RC workarea count higher than PLC workarea count -> Synchronization not possible 
  ERR_SYNC_WORKAREA_COUNT_RC_HIGHER_THAN_PLC := 19,

  
  /// END
  {warning 'ToDo: This is an internal error ID, which is not defined in SRCI specification'}
  
  
  
  
  /// Telegram control does not match the telegram state
  ERR_TELEGRAM_CONTROL_MISMATCH_TELEGRAM_STATE_0xA1 := 16#A1,  
  /// Initialization lost for unknown reason. See message log after reinitializing
  ERR_INIT_LOST_UNKNOWN_0xA2  := 16#A2,
  /// Telegram length does not match the length provided in the communication interface.
  ERR_TELEGRAM_LENGTH_MISMATCH_0xA3 := 16#A3,
  /// Incompatible major SRCI version
  ERR_SRCI_MAJOR_VERSION_INCOMPATIBLE_0xA4 := 16#A4,
  /// Lifesign timeout
  ERR_LIFESIGN_TIMEOUT_0xA5 := 16#A5,
  /// The selected optional cyclic data does not fit in the given telegram size
  ERR_CYCLIC_DATA_TOO_LARGE_0xA6 := 16#A6,
  /// The robot interface was reset after being initialized
  ERR_INTERFACE_WAS_RESET_AFTER_INIT_0xA7 := 16#A7,
  /// Telegram sequence timeout
  ERR_TELEGRAM_SEQ_TIMEOUT_0xA8 := 16#A8,
  /// The telegram number changed after initialization
  ERR_TELEGRAM_NO_CHANGED_AFTER_INIT_0xA9 := 16#A9,
  /// Invalid AxesGroupID
  ERR_AXESGROUP_ID_INVALID_0xAA := 16#AA,
  /// Telegram number is invalid. E.g. TwoSequences is only activated in one direction
  ERR_TELEGRAM_NUMBER_INVALID_0xAB := 16#AB,
  /// Telegram Number is not supported
  ERR_TELEGRAM_NUMBER_NOT_SUPPORTED_0xAC := 16#AC,
  /// Server Connection to the communication partner was lost
  ERR_SERVER_CONNECTION_LOST_0xAD := 16#AD,
  
  
  /// Table 5-103: Telegram and Initialization State 
  /// Initialization may fail due to several reasons, described in the following table. T he failure is
  /// signaled using the telegram state byte.
 

  /// 7.1 Table "A" – Command ErrorIDs 
  /// If an error related to the execution of a function block occurs, the function block returns an ErrorID
  /// to specify the error. The errors are stored in the PLC message buffer and are displayed on the
  /// function block outputs.
  /// In the PLC message buffer, they are dynamically arranged by the client to be displayed as follows:
  /// <Origin> <MessageType> <Command name> <Description>
  /// More information about the general message handling mechanism can be found in 5.5.11
  /// Diagnostics.
  /// The following table gives an overview over the existing ErrorIDs reported by commands and the
  /// corresponding description.

  /// ------------------------------------------------------
  /// CLIENT ErrorIDs
  /// ------------------------------------------------------

  /// Client Specified Velocity not valid
  /// Commands using the parameter "Velocity"
  ERR_VELOCITY_INVALID  := 16#8401,
  
  /// Client Specified Acceleration not valid
  /// Commands using the parameter "Acceleration"
  ERR_ACCELERATION_INVALID  := 16#8402,
  
  /// Client Specified Deceleration not valid
  /// Commands using the parameter "Deceleration"
  ERR_DECELERATION_INVALID  := 16#8403,
  
  /// Client Specified Jerk not valid
  /// Commands using the parameter "Jerk"
  ERR_JERK_INVALID  := 16#8404,
  
  /// Client Invalid parameter value - ConfigMode Elbow
  /// Commands using the parameter "ConfigMode"
  ERR_CONFIGMODE_ELBOW_INVALID  := 16#8405,
  
  /// Client Invalid parameter value - ConfigMode Shoulder
  /// Commands using the parameter "ConfigMode"
  ERR_CONFIGMODE_SHOULDER_INVALID  := 16#8406,
  
  /// Client Invalid parameter value - ConfigMode Wrist
  /// Commands using the parameter "ConfigMode"
  ERR_CONFIGMODE_WRIST_INVALID  := 16#8407,
  
  /// Client Invalid parameter value - TrajectoryMode
  /// Commands using the parameter "TrajectoryMode"
  ERR_TRAJECTORYMODE_INVALID  := 16#8409,
  
  /// Client Invalid parameter value - Override
  /// Commands using the parameter "Override"
  ERR_OVERRIDE_INVALID  := 16#8410,
  
  /// Client Invalid parameter value - AbortingMode.
  /// Only 0: Buffer / 1: Abort are valid.
  /// Commands using the parameter "AbortingMode"
  ERR_ABORTINGMODE_INVALID  := 16#8411,
  
  /// Client Invalid parameter value - ToolNo outside of
  /// the allowed range -1..254
  /// Commands using the parameter "ToolNo"
  ERR_TOOLNO_RANGE  := 16#8412,
  
  /// Client Invalid parameter value - ToolNo not
  /// available on RC
  /// Commands using the parameter "ToolNo"
  ERR_TOOLNO_UNAVAILABLE  := 16#8413,
  
  /// Client Invalid parameter value - FrameNo outside
  /// of the allowed range -1..254
  /// Commands using the parameter "FrameNo"
  ERR_FRAMENO_RANGE  := 16#8414,
  
  /// Client Invalid parameter value - FrameNo not
  /// available on RC
  /// Commands using the parameter "FrameNo"
  ERR_FRAMENO_UNAVAILABLE  := 16#8415,
  
  /// Client The array specified for AcyclicData exceeds
  /// the supported maximum length of 190 bytes
  /// Command "CallSubprogram"
  ERR_ACYCLICDATA_TOO_LARGE  := 16#8416,
  
  /// Client The array length specified for ReturnAcyclicData
  /// is not sufficient for the returned data. The data has been truncated
  /// Command "CallSubprogram"
  ERR_RETURNACYCLICDATA_TRUNCATED  := 16#8417,
  
  /// Client Invalid parameter value - LoadNo outside of
  /// the allowed range -1..254
  /// All commands
  ERR_LOADNO_RANGE  := 16#8418,
  
  /// Invalid parameter value - the requested ExportMode does not exist
  ERR_EXPORTMODE_NOT_EXIST := 16#8419,
  
  /// Invalid parameter value - the requested ExportName does not exist
  ERR_EXPORTNAME_NOT_EXIST := 16#8420,
  
  /// The given ExportName is already exist
  ERR_EXPORTNAME_ALREADY_EXISTS := 16#8421,
  
  /// No memory is left for data log
  ERR_DATALOG_NO_MEMORY_LEFT := 16#8422,
  
  /// An Error occurred during data loging . Message encludes Error ID
  ERR_DATALOG_ERROR_OCCURRED := 16#8425,
  
  /// Internal System Error "Undefined Step"
  ERR_INTERNAL_UNDEFINED_STEP := 16#8601,
  
  /// Client Specified ProcessingMode not defined
  /// Commands using the parameter "ProcessingMode"
  ERR_PROCESSINGMODE_NOT_DEFINED  := 16#8602,
  
  /// Client Specified ProcessingMode not allowed
  /// Commands using the parameter "ProcessingMode"
  ERR_PROCESSINGMODE_NOT_ALLOWED  := 16#8603,
  
  /// Client Specified Emitter ID not allowed
  /// Commands using the parameter "EmitterID"
  ERR_EMITTERID_NOT_ALLOWED := 16#8604,
  
  /// Client Specified Listener ID not allowed
  /// Commands using the parameter "ListenerID"
  ERR_LISTENERID_NOT_ALLOWED   := 16#8605,
  
  /// Client ProcessingMode or SequenceFlag changed during execution
  /// Commands using the parameter "ProcessingMode" or "SequenceFlag"
  ERR_PROCSEQFLAG_CHANGED  := 16#8609,
  
  /// Specified priority to high
  ERR_PRIORITY_TOO_LOW := 16#8610,

  /// Specified priority to low
  ERR_PRIORITY_TOO_HIGH := 16#8611,
  
  /// Client Commands are not Enabled (First Robot must be initialized)
  /// All commands
  ERR_COMMANDS_NOT_ENABLED  := 16#8612,
  
